(* IEC 61131-3 sources: veristc/veri-stc/tests/st-examples (part 4) *)

cond_a := LimitHigh(raw_110_a, 130);
cond_a := cond_a AND quality_a;
cond_a := cond_a AND (NOT bypass_a);
input_valid_a := InputValid(raw_110_a, 0, 1000);
cond_a := cond_a AND input_valid_a;
IF NOT input_valid_a THEN
    channel_fault_a := channel_fault_a + 1;
END_IF;
cond_b := LimitHigh(raw_110_b, 130);
cond_b := cond_b AND quality_b;
cond_b := cond_b AND (NOT bypass_b);
input_valid_b := InputValid(raw_110_b, 0, 1000);
cond_b := cond_b AND input_valid_b;
IF NOT input_valid_b THEN
    channel_fault_b := channel_fault_b + 1;
END_IF;
cond_c := LimitHigh(raw_110_c, 130);
cond_c := cond_c AND quality_c;
cond_c := cond_c AND (NOT bypass_c);
input_valid_c := InputValid(raw_110_c, 0, 1000);
cond_c := cond_c AND input_valid_c;
IF NOT input_valid_c THEN
    channel_fault_c := channel_fault_c + 1;
END_IF;
cond_d := LimitHigh(raw_110_d, 130);
cond_d := cond_d AND quality_d;
cond_d := cond_d AND (NOT bypass_d);
input_valid_d := InputValid(raw_110_d, 0, 1000);
cond_d := cond_d AND input_valid_d;
IF NOT input_valid_d THEN
    channel_fault_d := channel_fault_d + 1;
END_IF;
vote_ok := TwoOfFour(cond_a, cond_b, cond_c, cond_d);
IF cond_a <> cond_b THEN
    diagnosis_count := diagnosis_count + 1;
END_IF;
IF cond_c <> cond_d THEN
    diagnosis_count := diagnosis_count + 1;
END_IF;
IF NOT vote_ok THEN
    diagnosis_count := diagnosis_count + 1;
END_IF;
latch_a_110 := RS_Next(vote_ok, train_a_reset, latch_a_110);
IF latch_a_110 AND (NOT train_a_inhibit) THEN
    mask_a_13 := mask_a_13 + 64;
    trip_a := 0 < 1;
    scram_a := 0 < 1;
    breaker_a := 0 > 1;
    mfw_a := 0 < 1;
    alarm_a := 0 < 1;
END_IF;
latch_b_110 := RS_Next(vote_ok, train_b_reset, latch_b_110);
IF latch_b_110 AND (NOT train_b_inhibit) THEN
    mask_b_13 := mask_b_13 + 64;
    trip_b := 0 < 1;
    scram_b := 0 < 1;
    breaker_b := 0 > 1;
    mfw_b := 0 < 1;
    alarm_b := 0 < 1;
END_IF;
IF (raw_110_a > 130) AND (NOT cond_a) THEN
    channel_fault_a := channel_fault_a + 1;
END_IF;
IF (raw_110_b > 130) AND (NOT cond_b) THEN
    channel_fault_b := channel_fault_b + 1;
END_IF;
IF (raw_110_c > 130) AND (NOT cond_c) THEN
    channel_fault_c := channel_fault_c + 1;
END_IF;
IF (raw_110_d > 130) AND (NOT cond_d) THEN
    channel_fault_d := channel_fault_d + 1;
END_IF;
IF vote_ok AND train_a_inhibit THEN
    diagnosis_count := diagnosis_count + 1;
END_IF;
IF vote_ok AND train_b_inhibit THEN
    diagnosis_count := diagnosis_count + 1;
END_IF;

cond_a := LimitHigh(raw_111_a, 131);
cond_a := cond_a AND quality_a;
cond_a := cond_a AND (NOT bypass_a);
input_valid_a := InputValid(raw_111_a, 0, 1000);
cond_a := cond_a AND input_valid_a;
IF NOT input_valid_a THEN
    channel_fault_a := channel_fault_a + 1;
END_IF;
cond_b := LimitHigh(raw_111_b, 131);
cond_b := cond_b AND quality_b;
cond_b := cond_b AND (NOT bypass_b);
input_valid_b := InputValid(raw_111_b, 0, 1000);
cond_b := cond_b AND input_valid_b;
IF NOT input_valid_b THEN
    channel_fault_b := channel_fault_b + 1;
END_IF;
cond_c := LimitHigh(raw_111_c, 131);
cond_c := cond_c AND quality_c;
cond_c := cond_c AND (NOT bypass_c);
input_valid_c := InputValid(raw_111_c, 0, 1000);
cond_c := cond_c AND input_valid_c;
IF NOT input_valid_c THEN
    channel_fault_c := channel_fault_c + 1;
END_IF;
cond_d := LimitHigh(raw_111_d, 131);
cond_d := cond_d AND quality_d;
cond_d := cond_d AND (NOT bypass_d);
input_valid_d := InputValid(raw_111_d, 0, 1000);
cond_d := cond_d AND input_valid_d;
IF NOT input_valid_d THEN
    channel_fault_d := channel_fault_d + 1;
END_IF;
vote_ok := TwoOfFour(cond_a, cond_b, cond_c, cond_d);
IF cond_a <> cond_b THEN
    diagnosis_count := diagnosis_count + 1;
END_IF;
IF cond_c <> cond_d THEN
    diagnosis_count := diagnosis_count + 1;
END_IF;
IF NOT vote_ok THEN
    diagnosis_count := diagnosis_count + 1;
END_IF;
latch_a_111 := RS_Next(vote_ok, train_a_reset, latch_a_111);
IF latch_a_111 AND (NOT train_a_inhibit) THEN
    mask_a_13 := mask_a_13 + 128;
    trip_a := 0 < 1;
    scram_a := 0 < 1;
    breaker_a := 0 > 1;
    afw_a := 0 < 1;
    alarm_a := 0 < 1;
END_IF;
latch_b_111 := RS_Next(vote_ok, train_b_reset, latch_b_111);
IF latch_b_111 AND (NOT train_b_inhibit) THEN
    mask_b_13 := mask_b_13 + 128;
    trip_b := 0 < 1;
    scram_b := 0 < 1;
    breaker_b := 0 > 1;
    afw_b := 0 < 1;
    alarm_b := 0 < 1;
END_IF;
IF (raw_111_a > 131) AND (NOT cond_a) THEN
    channel_fault_a := channel_fault_a + 1;
END_IF;
IF (raw_111_b > 131) AND (NOT cond_b) THEN
    channel_fault_b := channel_fault_b + 1;
END_IF;
IF (raw_111_c > 131) AND (NOT cond_c) THEN
    channel_fault_c := channel_fault_c + 1;
END_IF;
IF (raw_111_d > 131) AND (NOT cond_d) THEN
    channel_fault_d := channel_fault_d + 1;
END_IF;
IF vote_ok AND train_a_inhibit THEN
    diagnosis_count := diagnosis_count + 1;
END_IF;
IF vote_ok AND train_b_inhibit THEN
    diagnosis_count := diagnosis_count + 1;
END_IF;

cond_a := LimitHigh(raw_112_a, 132);
cond_a := cond_a AND quality_a;
cond_a := cond_a AND (NOT bypass_a);
input_valid_a := InputValid(raw_112_a, 0, 1000);
cond_a := cond_a AND input_valid_a;
IF NOT input_valid_a THEN
    channel_fault_a := channel_fault_a + 1;
END_IF;
cond_b := LimitHigh(raw_112_b, 132);
cond_b := cond_b AND quality_b;
cond_b := cond_b AND (NOT bypass_b);
input_valid_b := InputValid(raw_112_b, 0, 1000);
cond_b := cond_b AND input_valid_b;
IF NOT input_valid_b THEN
    channel_fault_b := channel_fault_b + 1;
END_IF;
cond_c := LimitHigh(raw_112_c, 132);
cond_c := cond_c AND quality_c;
cond_c := cond_c AND (NOT bypass_c);
input_valid_c := InputValid(raw_112_c, 0, 1000);
cond_c := cond_c AND input_valid_c;
IF NOT input_valid_c THEN
    channel_fault_c := channel_fault_c + 1;
END_IF;
cond_d := LimitHigh(raw_112_d, 132);
cond_d := cond_d AND quality_d;
cond_d := cond_d AND (NOT bypass_d);
input_valid_d := InputValid(raw_112_d, 0, 1000);
cond_d := cond_d AND input_valid_d;
IF NOT input_valid_d THEN
    channel_fault_d := channel_fault_d + 1;
END_IF;
vote_ok := TwoOfFour(cond_a, cond_b, cond_c, cond_d);
IF cond_a <> cond_b THEN
    diagnosis_count := diagnosis_count + 1;
END_IF;
IF cond_c <> cond_d THEN
    diagnosis_count := diagnosis_count + 1;
END_IF;
IF NOT vote_ok THEN
    diagnosis_count := diagnosis_count + 1;
END_IF;
latch_a_112 := RS_Next(vote_ok, train_a_reset, latch_a_112);
IF latch_a_112 AND (NOT train_a_inhibit) THEN
    mask_a_14 := mask_a_14 + 1;
    trip_a := 0 < 1;
    scram_a := 0 < 1;
    breaker_a := 0 > 1;
    si_a := 0 < 1;
    alarm_a := 0 < 1;
END_IF;
latch_b_112 := RS_Next(vote_ok, train_b_reset, latch_b_112);
IF latch_b_112 AND (NOT train_b_inhibit) THEN
    mask_b_14 := mask_b_14 + 1;
    trip_b := 0 < 1;
    scram_b := 0 < 1;
    breaker_b := 0 > 1;
    si_b := 0 < 1;
    alarm_b := 0 < 1;
END_IF;
IF (raw_112_a > 132) AND (NOT cond_a) THEN
    channel_fault_a := channel_fault_a + 1;
END_IF;
IF (raw_112_b > 132) AND (NOT cond_b) THEN
    channel_fault_b := channel_fault_b + 1;
END_IF;
IF (raw_112_c > 132) AND (NOT cond_c) THEN
    channel_fault_c := channel_fault_c + 1;
END_IF;
IF (raw_112_d > 132) AND (NOT cond_d) THEN
    channel_fault_d := channel_fault_d + 1;
END_IF;
IF vote_ok AND train_a_inhibit THEN
    diagnosis_count := diagnosis_count + 1;
END_IF;
IF vote_ok AND train_b_inhibit THEN
    diagnosis_count := diagnosis_count + 1;
END_IF;

cond_a := LimitHigh(raw_113_a, 133);
cond_a := cond_a AND quality_a;
cond_a := cond_a AND (NOT bypass_a);
input_valid_a := InputValid(raw_113_a, 0, 1000);
cond_a := cond_a AND input_valid_a;
IF NOT input_valid_a THEN
    channel_fault_a := channel_fault_a + 1;
END_IF;
cond_b := LimitHigh(raw_113_b, 133);
cond_b := cond_b AND quality_b;
cond_b := cond_b AND (NOT bypass_b);
input_valid_b := InputValid(raw_113_b, 0, 1000);
cond_b := cond_b AND input_valid_b;
IF NOT input_valid_b THEN
    channel_fault_b := channel_fault_b + 1;
END_IF;
cond_c := LimitHigh(raw_113_c, 133);
cond_c := cond_c AND quality_c;
cond_c := cond_c AND (NOT bypass_c);
input_valid_c := InputValid(raw_113_c, 0, 1000);
cond_c := cond_c AND input_valid_c;
IF NOT input_valid_c THEN
    channel_fault_c := channel_fault_c + 1;
END_IF;
cond_d := LimitHigh(raw_113_d, 133);
cond_d := cond_d AND quality_d;
cond_d := cond_d AND (NOT bypass_d);
input_valid_d := InputValid(raw_113_d, 0, 1000);
cond_d := cond_d AND input_valid_d;
IF NOT input_valid_d THEN
    channel_fault_d := channel_fault_d + 1;
END_IF;
vote_ok := TwoOfFour(cond_a, cond_b, cond_c, cond_d);
IF cond_a <> cond_b THEN
    diagnosis_count := diagnosis_count + 1;
END_IF;
IF cond_c <> cond_d THEN
    diagnosis_count := diagnosis_count + 1;
END_IF;
IF NOT vote_ok THEN
    diagnosis_count := diagnosis_count + 1;
END_IF;
latch_a_113 := RS_Next(vote_ok, train_a_reset, latch_a_113);
IF latch_a_113 AND (NOT train_a_inhibit) THEN
    mask_a_14 := mask_a_14 + 2;
    trip_a := 0 < 1;
    scram_a := 0 < 1;
    breaker_a := 0 > 1;
    ci_a := 0 < 1;
    alarm_a := 0 < 1;
END_IF;
latch_b_113 := RS_Next(vote_ok, train_b_reset, latch_b_113);
IF latch_b_113 AND (NOT train_b_inhibit) THEN
    mask_b_14 := mask_b_14 + 2;
    trip_b := 0 < 1;
    scram_b := 0 < 1;
    breaker_b := 0 > 1;
    ci_b := 0 < 1;
    alarm_b := 0 < 1;
END_IF;
IF (raw_113_a > 133) AND (NOT cond_a) THEN
    channel_fault_a := channel_fault_a + 1;
END_IF;
IF (raw_113_b > 133) AND (NOT cond_b) THEN
    channel_fault_b := channel_fault_b + 1;
END_IF;
IF (raw_113_c > 133) AND (NOT cond_c) THEN
    channel_fault_c := channel_fault_c + 1;
END_IF;
IF (raw_113_d > 133) AND (NOT cond_d) THEN
    channel_fault_d := channel_fault_d + 1;
END_IF;
IF vote_ok AND train_a_inhibit THEN
    diagnosis_count := diagnosis_count + 1;
END_IF;
IF vote_ok AND train_b_inhibit THEN
    diagnosis_count := diagnosis_count + 1;
END_IF;

cond_a := LimitHigh(raw_114_a, 134);
cond_a := cond_a AND quality_a;
cond_a := cond_a AND (NOT bypass_a);
input_valid_a := InputValid(raw_114_a, 0, 1000);
cond_a := cond_a AND input_valid_a;
IF NOT input_valid_a THEN
    channel_fault_a := channel_fault_a + 1;
END_IF;
cond_b := LimitHigh(raw_114_b, 134);
cond_b := cond_b AND quality_b;
cond_b := cond_b AND (NOT bypass_b);
input_valid_b := InputValid(raw_114_b, 0, 1000);
cond_b := cond_b AND input_valid_b;
IF NOT input_valid_b THEN
    channel_fault_b := channel_fault_b + 1;
END_IF;
cond_c := LimitHigh(raw_114_c, 134);
cond_c := cond_c AND quality_c;
cond_c := cond_c AND (NOT bypass_c);
input_valid_c := InputValid(raw_114_c, 0, 1000);
cond_c := cond_c AND input_valid_c;
IF NOT input_valid_c THEN
    channel_fault_c := channel_fault_c + 1;
END_IF;
cond_d := LimitHigh(raw_114_d, 134);
cond_d := cond_d AND quality_d;
cond_d := cond_d AND (NOT bypass_d);
input_valid_d := InputValid(raw_114_d, 0, 1000);
cond_d := cond_d AND input_valid_d;
IF NOT input_valid_d THEN
    channel_fault_d := channel_fault_d + 1;
END_IF;
vote_ok := TwoOfFour(cond_a, cond_b, cond_c, cond_d);
IF cond_a <> cond_b THEN
    diagnosis_count := diagnosis_count + 1;
END_IF;
IF cond_c <> cond_d THEN
    diagnosis_count := diagnosis_count + 1;
END_IF;
IF NOT vote_ok THEN
    diagnosis_count := diagnosis_count + 1;
END_IF;
latch_a_114 := RS_Next(vote_ok, train_a_reset, latch_a_114);
IF latch_a_114 AND (NOT train_a_inhibit) THEN
    mask_a_14 := mask_a_14 + 4;
    trip_a := 0 < 1;
    scram_a := 0 < 1;
    breaker_a := 0 > 1;
    mfw_a := 0 < 1;
    alarm_a := 0 < 1;
END_IF;
latch_b_114 := RS_Next(vote_ok, train_b_reset, latch_b_114);
IF latch_b_114 AND (NOT train_b_inhibit) THEN
    mask_b_14 := mask_b_14 + 4;
    trip_b := 0 < 1;
    scram_b := 0 < 1;
    breaker_b := 0 > 1;
    mfw_b := 0 < 1;
    alarm_b := 0 < 1;
END_IF;
IF (raw_114_a > 134) AND (NOT cond_a) THEN
    channel_fault_a := channel_fault_a + 1;
END_IF;
IF (raw_114_b > 134) AND (NOT cond_b) THEN
    channel_fault_b := channel_fault_b + 1;
END_IF;
IF (raw_114_c > 134) AND (NOT cond_c) THEN
    channel_fault_c := channel_fault_c + 1;
END_IF;
IF (raw_114_d > 134) AND (NOT cond_d) THEN
    channel_fault_d := channel_fault_d + 1;
END_IF;
IF vote_ok AND train_a_inhibit THEN
    diagnosis_count := diagnosis_count + 1;
END_IF;
IF vote_ok AND train_b_inhibit THEN
    diagnosis_count := diagnosis_count + 1;
END_IF;

cond_a := LimitHigh(raw_115_a, 135);
cond_a := cond_a AND quality_a;
cond_a := cond_a AND (NOT bypass_a);
input_valid_a := InputValid(raw_115_a, 0, 1000);
cond_a := cond_a AND input_valid_a;
IF NOT input_valid_a THEN
    channel_fault_a := channel_fault_a + 1;
END_IF;
cond_b := LimitHigh(raw_115_b, 135);
cond_b := cond_b AND quality_b;
cond_b := cond_b AND (NOT bypass_b);
input_valid_b := InputValid(raw_115_b, 0, 1000);
cond_b := cond_b AND input_valid_b;
IF NOT input_valid_b THEN
    channel_fault_b := channel_fault_b + 1;
END_IF;
cond_c := LimitHigh(raw_115_c, 135);
cond_c := cond_c AND quality_c;
cond_c := cond_c AND (NOT bypass_c);
input_valid_c := InputValid(raw_115_c, 0, 1000);
cond_c := cond_c AND input_valid_c;
IF NOT input_valid_c THEN
    channel_fault_c := channel_fault_c + 1;
END_IF;
cond_d := LimitHigh(raw_115_d, 135);
cond_d := cond_d AND quality_d;
cond_d := cond_d AND (NOT bypass_d);
input_valid_d := InputValid(raw_115_d, 0, 1000);
cond_d := cond_d AND input_valid_d;
IF NOT input_valid_d THEN
    channel_fault_d := channel_fault_d + 1;
END_IF;
vote_ok := TwoOfFour(cond_a, cond_b, cond_c, cond_d);
IF cond_a <> cond_b THEN
    diagnosis_count := diagnosis_count + 1;
END_IF;
IF cond_c <> cond_d THEN
    diagnosis_count := diagnosis_count + 1;
END_IF;
IF NOT vote_ok THEN
    diagnosis_count := diagnosis_count + 1;
END_IF;
latch_a_115 := RS_Next(vote_ok, train_a_reset, latch_a_115);
IF latch_a_115 AND (NOT train_a_inhibit) THEN
    mask_a_14 := mask_a_14 + 8;
    trip_a := 0 < 1;
    scram_a := 0 < 1;
    breaker_a := 0 > 1;
    afw_a := 0 < 1;
    alarm_a := 0 < 1;
END_IF;
latch_b_115 := RS_Next(vote_ok, train_b_reset, latch_b_115);
IF latch_b_115 AND (NOT train_b_inhibit) THEN
    mask_b_14 := mask_b_14 + 8;
    trip_b := 0 < 1;
    scram_b := 0 < 1;
    breaker_b := 0 > 1;
    afw_b := 0 < 1;
    alarm_b := 0 < 1;
END_IF;
IF (raw_115_a > 135) AND (NOT cond_a) THEN
    channel_fault_a := channel_fault_a + 1;
END_IF;
IF (raw_115_b > 135) AND (NOT cond_b) THEN
    channel_fault_b := channel_fault_b + 1;
END_IF;
IF (raw_115_c > 135) AND (NOT cond_c) THEN
    channel_fault_c := channel_fault_c + 1;
END_IF;
IF (raw_115_d > 135) AND (NOT cond_d) THEN
    channel_fault_d := channel_fault_d + 1;
END_IF;
IF vote_ok AND train_a_inhibit THEN
    diagnosis_count := diagnosis_count + 1;
END_IF;
IF vote_ok AND train_b_inhibit THEN
    diagnosis_count := diagnosis_count + 1;
END_IF;

cond_a := LimitHigh(raw_116_a, 136);
cond_a := cond_a AND quality_a;
cond_a := cond_a AND (NOT bypass_a);
input_valid_a := InputValid(raw_116_a, 0, 1000);
cond_a := cond_a AND input_valid_a;
IF NOT input_valid_a THEN
    channel_fault_a := channel_fault_a + 1;
END_IF;
cond_b := LimitHigh(raw_116_b, 136);
cond_b := cond_b AND quality_b;
cond_b := cond_b AND (NOT bypass_b);
input_valid_b := InputValid(raw_116_b, 0, 1000);
cond_b := cond_b AND input_valid_b;
IF NOT input_valid_b THEN
    channel_fault_b := channel_fault_b + 1;
END_IF;
cond_c := LimitHigh(raw_116_c, 136);
cond_c := cond_c AND quality_c;
cond_c := cond_c AND (NOT bypass_c);
input_valid_c := InputValid(raw_116_c, 0, 1000);
cond_c := cond_c AND input_valid_c;
IF NOT input_valid_c THEN
    channel_fault_c := channel_fault_c + 1;
END_IF;
cond_d := LimitHigh(raw_116_d, 136);
cond_d := cond_d AND quality_d;
cond_d := cond_d AND (NOT bypass_d);
input_valid_d := InputValid(raw_116_d, 0, 1000);
cond_d := cond_d AND input_valid_d;
IF NOT input_valid_d THEN
    channel_fault_d := channel_fault_d + 1;
END_IF;
vote_ok := TwoOfFour(cond_a, cond_b, cond_c, cond_d);
IF cond_a <> cond_b THEN
    diagnosis_count := diagnosis_count + 1;
END_IF;
IF cond_c <> cond_d THEN
    diagnosis_count := diagnosis_count + 1;
END_IF;
IF NOT vote_ok THEN
    diagnosis_count := diagnosis_count + 1;
END_IF;
latch_a_116 := RS_Next(vote_ok, train_a_reset, latch_a_116);
IF latch_a_116 AND (NOT train_a_inhibit) THEN
    mask_a_14 := mask_a_14 + 16;
    trip_a := 0 < 1;
    scram_a := 0 < 1;
    breaker_a := 0 > 1;
    si_a := 0 < 1;
    alarm_a := 0 < 1;
END_IF;
latch_b_116 := RS_Next(vote_ok, train_b_reset, latch_b_116);
IF latch_b_116 AND (NOT train_b_inhibit) THEN
    mask_b_14 := mask_b_14 + 16;
    trip_b := 0 < 1;
    scram_b := 0 < 1;
    breaker_b := 0 > 1;
    si_b := 0 < 1;
    alarm_b := 0 < 1;
END_IF;
IF (raw_116_a > 136) AND (NOT cond_a) THEN
    channel_fault_a := channel_fault_a + 1;
END_IF;
IF (raw_116_b > 136) AND (NOT cond_b) THEN
    channel_fault_b := channel_fault_b + 1;
END_IF;
IF (raw_116_c > 136) AND (NOT cond_c) THEN
    channel_fault_c := channel_fault_c + 1;
END_IF;
IF (raw_116_d > 136) AND (NOT cond_d) THEN
    channel_fault_d := channel_fault_d + 1;
END_IF;
IF vote_ok AND train_a_inhibit THEN
    diagnosis_count := diagnosis_count + 1;
END_IF;
IF vote_ok AND train_b_inhibit THEN
    diagnosis_count := diagnosis_count + 1;
END_IF;

cond_a := LimitHigh(raw_117_a, 137);
cond_a := cond_a AND quality_a;
cond_a := cond_a AND (NOT bypass_a);
input_valid_a := InputValid(raw_117_a, 0, 1000);
cond_a := cond_a AND input_valid_a;
IF NOT input_valid_a THEN
    channel_fault_a := channel_fault_a + 1;
END_IF;
cond_b := LimitHigh(raw_117_b, 137);
cond_b := cond_b AND quality_b;
cond_b := cond_b AND (NOT bypass_b);
input_valid_b := InputValid(raw_117_b, 0, 1000);
cond_b := cond_b AND input_valid_b;
IF NOT input_valid_b THEN
    channel_fault_b := channel_fault_b + 1;
END_IF;
cond_c := LimitHigh(raw_117_c, 137);
cond_c := cond_c AND quality_c;
cond_c := cond_c AND (NOT bypass_c);
input_valid_c := InputValid(raw_117_c, 0, 1000);
cond_c := cond_c AND input_valid_c;
IF NOT input_valid_c THEN
    channel_fault_c := channel_fault_c + 1;
END_IF;
cond_d := LimitHigh(raw_117_d, 137);
cond_d := cond_d AND quality_d;
cond_d := cond_d AND (NOT bypass_d);
input_valid_d := InputValid(raw_117_d, 0, 1000);
cond_d := cond_d AND input_valid_d;
IF NOT input_valid_d THEN
    channel_fault_d := channel_fault_d + 1;
END_IF;
vote_ok := TwoOfFour(cond_a, cond_b, cond_c, cond_d);
IF cond_a <> cond_b THEN
    diagnosis_count := diagnosis_count + 1;
END_IF;
IF cond_c <> cond_d THEN
    diagnosis_count := diagnosis_count + 1;
END_IF;
IF NOT vote_ok THEN
    diagnosis_count := diagnosis_count + 1;
END_IF;
latch_a_117 := RS_Next(vote_ok, train_a_reset, latch_a_117);
IF latch_a_117 AND (NOT train_a_inhibit) THEN
    mask_a_14 := mask_a_14 + 32;
    trip_a := 0 < 1;
    scram_a := 0 < 1;
    breaker_a := 0 > 1;
    ci_a := 0 < 1;
    alarm_a := 0 < 1;
END_IF;
latch_b_117 := RS_Next(vote_ok, train_b_reset, latch_b_117);
IF latch_b_117 AND (NOT train_b_inhibit) THEN
    mask_b_14 := mask_b_14 + 32;
    trip_b := 0 < 1;
    scram_b := 0 < 1;
    breaker_b := 0 > 1;
    ci_b := 0 < 1;
    alarm_b := 0 < 1;
END_IF;
IF (raw_117_a > 137) AND (NOT cond_a) THEN
    channel_fault_a := channel_fault_a + 1;
END_IF;
IF (raw_117_b > 137) AND (NOT cond_b) THEN
    channel_fault_b := channel_fault_b + 1;
END_IF;
IF (raw_117_c > 137) AND (NOT cond_c) THEN
    channel_fault_c := channel_fault_c + 1;
END_IF;
IF (raw_117_d > 137) AND (NOT cond_d) THEN
    channel_fault_d := channel_fault_d + 1;
END_IF;
IF vote_ok AND train_a_inhibit THEN
    diagnosis_count := diagnosis_count + 1;
END_IF;
IF vote_ok AND train_b_inhibit THEN
    diagnosis_count := diagnosis_count + 1;
END_IF;

cond_a := LimitHigh(raw_118_a, 138);
cond_a := cond_a AND quality_a;
cond_a := cond_a AND (NOT bypass_a);
input_valid_a := InputValid(raw_118_a, 0, 1000);
cond_a := cond_a AND input_valid_a;
IF NOT input_valid_a THEN
    channel_fault_a := channel_fault_a + 1;
END_IF;
cond_b := LimitHigh(raw_118_b, 138);
cond_b := cond_b AND quality_b;
cond_b := cond_b AND (NOT bypass_b);
input_valid_b := InputValid(raw_118_b, 0, 1000);
cond_b := cond_b AND input_valid_b;
IF NOT input_valid_b THEN
    channel_fault_b := channel_fault_b + 1;
END_IF;
cond_c := LimitHigh(raw_118_c, 138);
cond_c := cond_c AND quality_c;
cond_c := cond_c AND (NOT bypass_c);
input_valid_c := InputValid(raw_118_c, 0, 1000);
cond_c := cond_c AND input_valid_c;
IF NOT input_valid_c THEN
    channel_fault_c := channel_fault_c + 1;
END_IF;
cond_d := LimitHigh(raw_118_d, 138);
cond_d := cond_d AND quality_d;
cond_d := cond_d AND (NOT bypass_d);
input_valid_d := InputValid(raw_118_d, 0, 1000);
cond_d := cond_d AND input_valid_d;
IF NOT input_valid_d THEN
    channel_fault_d := channel_fault_d + 1;
END_IF;
vote_ok := TwoOfFour(cond_a, cond_b, cond_c, cond_d);
IF cond_a <> cond_b THEN
    diagnosis_count := diagnosis_count + 1;
END_IF;
IF cond_c <> cond_d THEN
    diagnosis_count := diagnosis_count + 1;
END_IF;
IF NOT vote_ok THEN
    diagnosis_count := diagnosis_count + 1;
END_IF;
latch_a_118 := RS_Next(vote_ok, train_a_reset, latch_a_118);
IF latch_a_118 AND (NOT train_a_inhibit) THEN
    mask_a_14 := mask_a_14 + 64;
    trip_a := 0 < 1;
    scram_a := 0 < 1;
    breaker_a := 0 > 1;
    mfw_a := 0 < 1;
    alarm_a := 0 < 1;
END_IF;
latch_b_118 := RS_Next(vote_ok, train_b_reset, latch_b_118);
IF latch_b_118 AND (NOT train_b_inhibit) THEN
    mask_b_14 := mask_b_14 + 64;
    trip_b := 0 < 1;
    scram_b := 0 < 1;
    breaker_b := 0 > 1;
    mfw_b := 0 < 1;
    alarm_b := 0 < 1;
END_IF;
IF (raw_118_a > 138) AND (NOT cond_a) THEN
    channel_fault_a := channel_fault_a + 1;
END_IF;
IF (raw_118_b > 138) AND (NOT cond_b) THEN
    channel_fault_b := channel_fault_b + 1;
END_IF;
IF (raw_118_c > 138) AND (NOT cond_c) THEN
    channel_fault_c := channel_fault_c + 1;
END_IF;
IF (raw_118_d > 138) AND (NOT cond_d) THEN
    channel_fault_d := channel_fault_d + 1;
END_IF;
IF vote_ok AND train_a_inhibit THEN
    diagnosis_count := diagnosis_count + 1;
END_IF;
IF vote_ok AND train_b_inhibit THEN
    diagnosis_count := diagnosis_count + 1;
END_IF;

cond_a := LimitHigh(raw_119_a, 139);
cond_a := cond_a AND quality_a;
cond_a := cond_a AND (NOT bypass_a);
input_valid_a := InputValid(raw_119_a, 0, 1000);
cond_a := cond_a AND input_valid_a;
IF NOT input_valid_a THEN
    channel_fault_a := channel_fault_a + 1;
END_IF;
cond_b := LimitHigh(raw_119_b, 139);
cond_b := cond_b AND quality_b;
cond_b := cond_b AND (NOT bypass_b);
input_valid_b := InputValid(raw_119_b, 0, 1000);
cond_b := cond_b AND input_valid_b;
IF NOT input_valid_b THEN
    channel_fault_b := channel_fault_b + 1;
END_IF;
cond_c := LimitHigh(raw_119_c, 139);
cond_c := cond_c AND quality_c;
cond_c := cond_c AND (NOT bypass_c);
input_valid_c := InputValid(raw_119_c, 0, 1000);
cond_c := cond_c AND input_valid_c;
IF NOT input_valid_c THEN
    channel_fault_c := channel_fault_c + 1;
END_IF;
cond_d := LimitHigh(raw_119_d, 139);
cond_d := cond_d AND quality_d;
cond_d := cond_d AND (NOT bypass_d);
input_valid_d := InputValid(raw_119_d, 0, 1000);
cond_d := cond_d AND input_valid_d;
IF NOT input_valid_d THEN
    channel_fault_d := channel_fault_d + 1;
END_IF;
vote_ok := TwoOfFour(cond_a, cond_b, cond_c, cond_d);
IF cond_a <> cond_b THEN
    diagnosis_count := diagnosis_count + 1;
END_IF;
IF cond_c <> cond_d THEN
    diagnosis_count := diagnosis_count + 1;
END_IF;
IF NOT vote_ok THEN
    diagnosis_count := diagnosis_count + 1;
END_IF;
latch_a_119 := RS_Next(vote_ok, train_a_reset, latch_a_119);
IF latch_a_119 AND (NOT train_a_inhibit) THEN
    mask_a_14 := mask_a_14 + 128;
    trip_a := 0 < 1;
    scram_a := 0 < 1;
    breaker_a := 0 > 1;
    afw_a := 0 < 1;
    alarm_a := 0 < 1;
END_IF;
latch_b_119 := RS_Next(vote_ok, train_b_reset, latch_b_119);
IF latch_b_119 AND (NOT train_b_inhibit) THEN
    mask_b_14 := mask_b_14 + 128;
    trip_b := 0 < 1;
    scram_b := 0 < 1;
    breaker_b := 0 > 1;
    afw_b := 0 < 1;
    alarm_b := 0 < 1;
END_IF;
IF (raw_119_a > 139) AND (NOT cond_a) THEN
    channel_fault_a := channel_fault_a + 1;
END_IF;
IF (raw_119_b > 139) AND (NOT cond_b) THEN
    channel_fault_b := channel_fault_b + 1;
END_IF;
IF (raw_119_c > 139) AND (NOT cond_c) THEN
    channel_fault_c := channel_fault_c + 1;
END_IF;
IF (raw_119_d > 139) AND (NOT cond_d) THEN
    channel_fault_d := channel_fault_d + 1;
END_IF;
IF vote_ok AND train_a_inhibit THEN
    diagnosis_count := diagnosis_count + 1;
END_IF;
IF vote_ok AND train_b_inhibit THEN
    diagnosis_count := diagnosis_count + 1;
END_IF;

cond_a := LimitHigh(raw_120_a, 100);
cond_a := cond_a AND quality_a;
cond_a := cond_a AND (NOT bypass_a);
input_valid_a := InputValid(raw_120_a, 0, 1000);
cond_a := cond_a AND input_valid_a;
IF NOT input_valid_a THEN
    channel_fault_a := channel_fault_a + 1;
END_IF;
cond_b := LimitHigh(raw_120_b, 100);
cond_b := cond_b AND quality_b;
cond_b := cond_b AND (NOT bypass_b);
input_valid_b := InputValid(raw_120_b, 0, 1000);
cond_b := cond_b AND input_valid_b;
IF NOT input_valid_b THEN
    channel_fault_b := channel_fault_b + 1;
END_IF;
cond_c := LimitHigh(raw_120_c, 100);
cond_c := cond_c AND quality_c;
cond_c := cond_c AND (NOT bypass_c);
input_valid_c := InputValid(raw_120_c, 0, 1000);
cond_c := cond_c AND input_valid_c;
IF NOT input_valid_c THEN
    channel_fault_c := channel_fault_c + 1;
END_IF;
cond_d := LimitHigh(raw_120_d, 100);
cond_d := cond_d AND quality_d;
cond_d := cond_d AND (NOT bypass_d);
input_valid_d := InputValid(raw_120_d, 0, 1000);
cond_d := cond_d AND input_valid_d;
IF NOT input_valid_d THEN
    channel_fault_d := channel_fault_d + 1;
END_IF;
vote_ok := TwoOfFour(cond_a, cond_b, cond_c, cond_d);
IF cond_a <> cond_b THEN
    diagnosis_count := diagnosis_count + 1;
END_IF;
IF cond_c <> cond_d THEN
    diagnosis_count := diagnosis_count + 1;
END_IF;
IF NOT vote_ok THEN
    diagnosis_count := diagnosis_count + 1;
END_IF;
latch_a_120 := RS_Next(vote_ok, train_a_reset, latch_a_120);
IF latch_a_120 AND (NOT train_a_inhibit) THEN
    mask_a_15 := mask_a_15 + 1;
    trip_a := 0 < 1;
    scram_a := 0 < 1;
    breaker_a := 0 > 1;
    si_a := 0 < 1;
    alarm_a := 0 < 1;
END_IF;
latch_b_120 := RS_Next(vote_ok, train_b_reset, latch_b_120);
IF latch_b_120 AND (NOT train_b_inhibit) THEN
    mask_b_15 := mask_b_15 + 1;
    trip_b := 0 < 1;
    scram_b := 0 < 1;
    breaker_b := 0 > 1;
    si_b := 0 < 1;
    alarm_b := 0 < 1;
END_IF;
IF (raw_120_a > 100) AND (NOT cond_a) THEN
    channel_fault_a := channel_fault_a + 1;
END_IF;
IF (raw_120_b > 100) AND (NOT cond_b) THEN
    channel_fault_b := channel_fault_b + 1;
END_IF;
IF (raw_120_c > 100) AND (NOT cond_c) THEN
    channel_fault_c := channel_fault_c + 1;
END_IF;
IF (raw_120_d > 100) AND (NOT cond_d) THEN
    channel_fault_d := channel_fault_d + 1;
END_IF;
IF vote_ok AND train_a_inhibit THEN
    diagnosis_count := diagnosis_count + 1;
END_IF;
IF vote_ok AND train_b_inhibit THEN
    diagnosis_count := diagnosis_count + 1;
END_IF;

cond_a := LimitHigh(raw_121_a, 101);
cond_a := cond_a AND quality_a;
cond_a := cond_a AND (NOT bypass_a);
input_valid_a := InputValid(raw_121_a, 0, 1000);
cond_a := cond_a AND input_valid_a;
IF NOT input_valid_a THEN
    channel_fault_a := channel_fault_a + 1;
END_IF;
cond_b := LimitHigh(raw_121_b, 101);
cond_b := cond_b AND quality_b;
cond_b := cond_b AND (NOT bypass_b);
input_valid_b := InputValid(raw_121_b, 0, 1000);
cond_b := cond_b AND input_valid_b;
IF NOT input_valid_b THEN
    channel_fault_b := channel_fault_b + 1;
END_IF;
cond_c := LimitHigh(raw_121_c, 101);
cond_c := cond_c AND quality_c;
cond_c := cond_c AND (NOT bypass_c);
input_valid_c := InputValid(raw_121_c, 0, 1000);
cond_c := cond_c AND input_valid_c;
IF NOT input_valid_c THEN
    channel_fault_c := channel_fault_c + 1;
END_IF;
cond_d := LimitHigh(raw_121_d, 101);
cond_d := cond_d AND quality_d;
cond_d := cond_d AND (NOT bypass_d);
input_valid_d := InputValid(raw_121_d, 0, 1000);
cond_d := cond_d AND input_valid_d;
IF NOT input_valid_d THEN
    channel_fault_d := channel_fault_d + 1;
END_IF;
vote_ok := TwoOfFour(cond_a, cond_b, cond_c, cond_d);
IF cond_a <> cond_b THEN
    diagnosis_count := diagnosis_count + 1;
END_IF;
IF cond_c <> cond_d THEN
    diagnosis_count := diagnosis_count + 1;
END_IF;
IF NOT vote_ok THEN
    diagnosis_count := diagnosis_count + 1;
END_IF;
latch_a_121 := RS_Next(vote_ok, train_a_reset, latch_a_121);
IF latch_a_121 AND (NOT train_a_inhibit) THEN
    mask_a_15 := mask_a_15 + 2;
    trip_a := 0 < 1;
    scram_a := 0 < 1;
    breaker_a := 0 > 1;
    ci_a := 0 < 1;
    alarm_a := 0 < 1;
END_IF;
latch_b_121 := RS_Next(vote_ok, train_b_reset, latch_b_121);
IF latch_b_121 AND (NOT train_b_inhibit) THEN
    mask_b_15 := mask_b_15 + 2;
    trip_b := 0 < 1;
    scram_b := 0 < 1;
    breaker_b := 0 > 1;
    ci_b := 0 < 1;
    alarm_b := 0 < 1;
END_IF;
IF (raw_121_a > 101) AND (NOT cond_a) THEN
    channel_fault_a := channel_fault_a + 1;
END_IF;
IF (raw_121_b > 101) AND (NOT cond_b) THEN
    channel_fault_b := channel_fault_b + 1;
END_IF;
IF (raw_121_c > 101) AND (NOT cond_c) THEN
    channel_fault_c := channel_fault_c + 1;
END_IF;
IF (raw_121_d > 101) AND (NOT cond_d) THEN
    channel_fault_d := channel_fault_d + 1;
END_IF;
IF vote_ok AND train_a_inhibit THEN
    diagnosis_count := diagnosis_count + 1;
END_IF;
IF vote_ok AND train_b_inhibit THEN
    diagnosis_count := diagnosis_count + 1;
END_IF;

cond_a := LimitHigh(raw_122_a, 102);
cond_a := cond_a AND quality_a;
cond_a := cond_a AND (NOT bypass_a);
input_valid_a := InputValid(raw_122_a, 0, 1000);
cond_a := cond_a AND input_valid_a;
IF NOT input_valid_a THEN
    channel_fault_a := channel_fault_a + 1;
END_IF;
cond_b := LimitHigh(raw_122_b, 102);
cond_b := cond_b AND quality_b;
cond_b := cond_b AND (NOT bypass_b);
input_valid_b := InputValid(raw_122_b, 0, 1000);
cond_b := cond_b AND input_valid_b;
IF NOT input_valid_b THEN
    channel_fault_b := channel_fault_b + 1;
END_IF;
cond_c := LimitHigh(raw_122_c, 102);
cond_c := cond_c AND quality_c;
cond_c := cond_c AND (NOT bypass_c);
input_valid_c := InputValid(raw_122_c, 0, 1000);
cond_c := cond_c AND input_valid_c;
IF NOT input_valid_c THEN
    channel_fault_c := channel_fault_c + 1;
END_IF;
cond_d := LimitHigh(raw_122_d, 102);
cond_d := cond_d AND quality_d;
cond_d := cond_d AND (NOT bypass_d);
input_valid_d := InputValid(raw_122_d, 0, 1000);
cond_d := cond_d AND input_valid_d;
IF NOT input_valid_d THEN
    channel_fault_d := channel_fault_d + 1;
END_IF;
vote_ok := TwoOfFour(cond_a, cond_b, cond_c, cond_d);
IF cond_a <> cond_b THEN
    diagnosis_count := diagnosis_count + 1;
END_IF;
IF cond_c <> cond_d THEN
    diagnosis_count := diagnosis_count + 1;
END_IF;
IF NOT vote_ok THEN
    diagnosis_count := diagnosis_count + 1;
END_IF;
latch_a_122 := RS_Next(vote_ok, train_a_reset, latch_a_122);
IF latch_a_122 AND (NOT train_a_inhibit) THEN
    mask_a_15 := mask_a_15 + 4;
    trip_a := 0 < 1;
    scram_a := 0 < 1;
    breaker_a := 0 > 1;
    mfw_a := 0 < 1;
    alarm_a := 0 < 1;
END_IF;
latch_b_122 := RS_Next(vote_ok, train_b_reset, latch_b_122);
IF latch_b_122 AND (NOT train_b_inhibit) THEN
    mask_b_15 := mask_b_15 + 4;
    trip_b := 0 < 1;
    scram_b := 0 < 1;
    breaker_b := 0 > 1;
    mfw_b := 0 < 1;
    alarm_b := 0 < 1;
END_IF;
IF (raw_122_a > 102) AND (NOT cond_a) THEN
    channel_fault_a := channel_fault_a + 1;
END_IF;
IF (raw_122_b > 102) AND (NOT cond_b) THEN
    channel_fault_b := channel_fault_b + 1;
END_IF;
IF (raw_122_c > 102) AND (NOT cond_c) THEN
    channel_fault_c := channel_fault_c + 1;
END_IF;
IF (raw_122_d > 102) AND (NOT cond_d) THEN
    channel_fault_d := channel_fault_d + 1;
END_IF;
IF vote_ok AND train_a_inhibit THEN
    diagnosis_count := diagnosis_count + 1;
END_IF;
IF vote_ok AND train_b_inhibit THEN
    diagnosis_count := diagnosis_count + 1;
END_IF;

cond_a := LimitHigh(raw_123_a, 103);
cond_a := cond_a AND quality_a;
cond_a := cond_a AND (NOT bypass_a);
input_valid_a := InputValid(raw_123_a, 0, 1000);
cond_a := cond_a AND input_valid_a;
IF NOT input_valid_a THEN
    channel_fault_a := channel_fault_a + 1;
END_IF;
cond_b := LimitHigh(raw_123_b, 103);
cond_b := cond_b AND quality_b;
cond_b := cond_b AND (NOT bypass_b);
input_valid_b := InputValid(raw_123_b, 0, 1000);
cond_b := cond_b AND input_valid_b;
IF NOT input_valid_b THEN
    channel_fault_b := channel_fault_b + 1;
END_IF;
cond_c := LimitHigh(raw_123_c, 103);
cond_c := cond_c AND quality_c;
cond_c := cond_c AND (NOT bypass_c);
input_valid_c := InputValid(raw_123_c, 0, 1000);
cond_c := cond_c AND input_valid_c;
IF NOT input_valid_c THEN
    channel_fault_c := channel_fault_c + 1;
END_IF;
cond_d := LimitHigh(raw_123_d, 103);
cond_d := cond_d AND quality_d;
cond_d := cond_d AND (NOT bypass_d);
input_valid_d := InputValid(raw_123_d, 0, 1000);
cond_d := cond_d AND input_valid_d;
IF NOT input_valid_d THEN
    channel_fault_d := channel_fault_d + 1;
END_IF;
vote_ok := TwoOfFour(cond_a, cond_b, cond_c, cond_d);
IF cond_a <> cond_b THEN
    diagnosis_count := diagnosis_count + 1;
END_IF;
IF cond_c <> cond_d THEN
    diagnosis_count := diagnosis_count + 1;
END_IF;
IF NOT vote_ok THEN
    diagnosis_count := diagnosis_count + 1;
END_IF;
latch_a_123 := RS_Next(vote_ok, train_a_reset, latch_a_123);
IF latch_a_123 AND (NOT train_a_inhibit) THEN
    mask_a_15 := mask_a_15 + 8;
    trip_a := 0 < 1;
    scram_a := 0 < 1;
    breaker_a := 0 > 1;
    afw_a := 0 < 1;
    alarm_a := 0 < 1;
END_IF;
latch_b_123 := RS_Next(vote_ok, train_b_reset, latch_b_123);
IF latch_b_123 AND (NOT train_b_inhibit) THEN
    mask_b_15 := mask_b_15 + 8;
    trip_b := 0 < 1;
    scram_b := 0 < 1;
    breaker_b := 0 > 1;
    afw_b := 0 < 1;
    alarm_b := 0 < 1;
END_IF;
IF (raw_123_a > 103) AND (NOT cond_a) THEN
    channel_fault_a := channel_fault_a + 1;
END_IF;
IF (raw_123_b > 103) AND (NOT cond_b) THEN
    channel_fault_b := channel_fault_b + 1;
END_IF;
IF (raw_123_c > 103) AND (NOT cond_c) THEN
    channel_fault_c := channel_fault_c + 1;
END_IF;
IF (raw_123_d > 103) AND (NOT cond_d) THEN
    channel_fault_d := channel_fault_d + 1;
END_IF;
IF vote_ok AND train_a_inhibit THEN
    diagnosis_count := diagnosis_count + 1;
END_IF;
IF vote_ok AND train_b_inhibit THEN
    diagnosis_count := diagnosis_count + 1;
END_IF;

cond_a := LimitHigh(raw_124_a, 104);
cond_a := cond_a AND quality_a;
cond_a := cond_a AND (NOT bypass_a);
input_valid_a := InputValid(raw_124_a, 0, 1000);
cond_a := cond_a AND input_valid_a;
IF NOT input_valid_a THEN
    channel_fault_a := channel_fault_a + 1;
END_IF;
cond_b := LimitHigh(raw_124_b, 104);
cond_b := cond_b AND quality_b;
cond_b := cond_b AND (NOT bypass_b);
input_valid_b := InputValid(raw_124_b, 0, 1000);
cond_b := cond_b AND input_valid_b;
IF NOT input_valid_b THEN
    channel_fault_b := channel_fault_b + 1;
END_IF;
cond_c := LimitHigh(raw_124_c, 104);
cond_c := cond_c AND quality_c;
cond_c := cond_c AND (NOT bypass_c);
input_valid_c := InputValid(raw_124_c, 0, 1000);
cond_c := cond_c AND input_valid_c;
IF NOT input_valid_c THEN
    channel_fault_c := channel_fault_c + 1;
END_IF;
cond_d := LimitHigh(raw_124_d, 104);
cond_d := cond_d AND quality_d;
cond_d := cond_d AND (NOT bypass_d);
input_valid_d := InputValid(raw_124_d, 0, 1000);
cond_d := cond_d AND input_valid_d;
IF NOT input_valid_d THEN
    channel_fault_d := channel_fault_d + 1;
END_IF;
vote_ok := TwoOfFour(cond_a, cond_b, cond_c, cond_d);
IF cond_a <> cond_b THEN
    diagnosis_count := diagnosis_count + 1;
END_IF;
IF cond_c <> cond_d THEN
    diagnosis_count := diagnosis_count + 1;
END_IF;
IF NOT vote_ok THEN
    diagnosis_count := diagnosis_count + 1;
END_IF;
latch_a_124 := RS_Next(vote_ok, train_a_reset, latch_a_124);
IF latch_a_124 AND (NOT train_a_inhibit) THEN
    mask_a_15 := mask_a_15 + 16;
    trip_a := 0 < 1;
    scram_a := 0 < 1;
    breaker_a := 0 > 1;
    si_a := 0 < 1;
    alarm_a := 0 < 1;
END_IF;
latch_b_124 := RS_Next(vote_ok, train_b_reset, latch_b_124);
IF latch_b_124 AND (NOT train_b_inhibit) THEN
    mask_b_15 := mask_b_15 + 16;
    trip_b := 0 < 1;
    scram_b := 0 < 1;
    breaker_b := 0 > 1;
    si_b := 0 < 1;
    alarm_b := 0 < 1;
END_IF;
IF (raw_124_a > 104) AND (NOT cond_a) THEN
    channel_fault_a := channel_fault_a + 1;
END_IF;
IF (raw_124_b > 104) AND (NOT cond_b) THEN
    channel_fault_b := channel_fault_b + 1;
END_IF;
IF (raw_124_c > 104) AND (NOT cond_c) THEN
    channel_fault_c := channel_fault_c + 1;
END_IF;
IF (raw_124_d > 104) AND (NOT cond_d) THEN
    channel_fault_d := channel_fault_d + 1;
END_IF;
IF vote_ok AND train_a_inhibit THEN
    diagnosis_count := diagnosis_count + 1;
END_IF;
IF vote_ok AND train_b_inhibit THEN
    diagnosis_count := diagnosis_count + 1;
END_IF;

cond_a := LimitHigh(raw_125_a, 105);
cond_a := cond_a AND quality_a;
cond_a := cond_a AND (NOT bypass_a);
input_valid_a := InputValid(raw_125_a, 0, 1000);
cond_a := cond_a AND input_valid_a;
IF NOT input_valid_a THEN
    channel_fault_a := channel_fault_a + 1;
END_IF;
cond_b := LimitHigh(raw_125_b, 105);
cond_b := cond_b AND quality_b;
cond_b := cond_b AND (NOT bypass_b);
input_valid_b := InputValid(raw_125_b, 0, 1000);
cond_b := cond_b AND input_valid_b;
IF NOT input_valid_b THEN
    channel_fault_b := channel_fault_b + 1;
END_IF;
cond_c := LimitHigh(raw_125_c, 105);
cond_c := cond_c AND quality_c;
cond_c := cond_c AND (NOT bypass_c);
input_valid_c := InputValid(raw_125_c, 0, 1000);
cond_c := cond_c AND input_valid_c;
IF NOT input_valid_c THEN
    channel_fault_c := channel_fault_c + 1;
END_IF;
cond_d := LimitHigh(raw_125_d, 105);
cond_d := cond_d AND quality_d;
cond_d := cond_d AND (NOT bypass_d);
input_valid_d := InputValid(raw_125_d, 0, 1000);
cond_d := cond_d AND input_valid_d;
IF NOT input_valid_d THEN
    channel_fault_d := channel_fault_d + 1;
END_IF;
vote_ok := TwoOfFour(cond_a, cond_b, cond_c, cond_d);
IF cond_a <> cond_b THEN
    diagnosis_count := diagnosis_count + 1;
END_IF;
IF cond_c <> cond_d THEN
    diagnosis_count := diagnosis_count + 1;
END_IF;
IF NOT vote_ok THEN
    diagnosis_count := diagnosis_count + 1;
END_IF;
latch_a_125 := RS_Next(vote_ok, train_a_reset, latch_a_125);
IF latch_a_125 AND (NOT train_a_inhibit) THEN
    mask_a_15 := mask_a_15 + 32;
    trip_a := 0 < 1;
    scram_a := 0 < 1;
    breaker_a := 0 > 1;
    ci_a := 0 < 1;
    alarm_a := 0 < 1;
END_IF;
latch_b_125 := RS_Next(vote_ok, train_b_reset, latch_b_125);
IF latch_b_125 AND (NOT train_b_inhibit) THEN
    mask_b_15 := mask_b_15 + 32;
    trip_b := 0 < 1;
    scram_b := 0 < 1;
    breaker_b := 0 > 1;
    ci_b := 0 < 1;
    alarm_b := 0 < 1;
END_IF;
IF (raw_125_a > 105) AND (NOT cond_a) THEN
    channel_fault_a := channel_fault_a + 1;
END_IF;
IF (raw_125_b > 105) AND (NOT cond_b) THEN
    channel_fault_b := channel_fault_b + 1;
END_IF;
IF (raw_125_c > 105) AND (NOT cond_c) THEN
    channel_fault_c := channel_fault_c + 1;
END_IF;
IF (raw_125_d > 105) AND (NOT cond_d) THEN
    channel_fault_d := channel_fault_d + 1;
END_IF;
IF vote_ok AND train_a_inhibit THEN
    diagnosis_count := diagnosis_count + 1;
END_IF;
IF vote_ok AND train_b_inhibit THEN
    diagnosis_count := diagnosis_count + 1;
END_IF;

cond_a := LimitHigh(raw_126_a, 106);
cond_a := cond_a AND quality_a;
cond_a := cond_a AND (NOT bypass_a);
input_valid_a := InputValid(raw_126_a, 0, 1000);
cond_a := cond_a AND input_valid_a;
IF NOT input_valid_a THEN
    channel_fault_a := channel_fault_a + 1;
END_IF;
cond_b := LimitHigh(raw_126_b, 106);
cond_b := cond_b AND quality_b;
cond_b := cond_b AND (NOT bypass_b);
input_valid_b := InputValid(raw_126_b, 0, 1000);
cond_b := cond_b AND input_valid_b;
IF NOT input_valid_b THEN
    channel_fault_b := channel_fault_b + 1;
END_IF;
cond_c := LimitHigh(raw_126_c, 106);
cond_c := cond_c AND quality_c;
cond_c := cond_c AND (NOT bypass_c);
input_valid_c := InputValid(raw_126_c, 0, 1000);
cond_c := cond_c AND input_valid_c;
IF NOT input_valid_c THEN
    channel_fault_c := channel_fault_c + 1;
END_IF;
cond_d := LimitHigh(raw_126_d, 106);
cond_d := cond_d AND quality_d;
cond_d := cond_d AND (NOT bypass_d);
input_valid_d := InputValid(raw_126_d, 0, 1000);
cond_d := cond_d AND input_valid_d;
IF NOT input_valid_d THEN
    channel_fault_d := channel_fault_d + 1;
END_IF;
vote_ok := TwoOfFour(cond_a, cond_b, cond_c, cond_d);
IF cond_a <> cond_b THEN
    diagnosis_count := diagnosis_count + 1;
END_IF;
IF cond_c <> cond_d THEN
    diagnosis_count := diagnosis_count + 1;
END_IF;
IF NOT vote_ok THEN
    diagnosis_count := diagnosis_count + 1;
END_IF;
latch_a_126 := RS_Next(vote_ok, train_a_reset, latch_a_126);
IF latch_a_126 AND (NOT train_a_inhibit) THEN
    mask_a_15 := mask_a_15 + 64;
    trip_a := 0 < 1;
    scram_a := 0 < 1;
    breaker_a := 0 > 1;
    mfw_a := 0 < 1;
    alarm_a := 0 < 1;
END_IF;
latch_b_126 := RS_Next(vote_ok, train_b_reset, latch_b_126);
IF latch_b_126 AND (NOT train_b_inhibit) THEN
    mask_b_15 := mask_b_15 + 64;
    trip_b := 0 < 1;
    scram_b := 0 < 1;
    breaker_b := 0 > 1;
    mfw_b := 0 < 1;
    alarm_b := 0 < 1;
END_IF;
IF (raw_126_a > 106) AND (NOT cond_a) THEN
    channel_fault_a := channel_fault_a + 1;
END_IF;
IF (raw_126_b > 106) AND (NOT cond_b) THEN
    channel_fault_b := channel_fault_b + 1;
END_IF;
IF (raw_126_c > 106) AND (NOT cond_c) THEN
    channel_fault_c := channel_fault_c + 1;
END_IF;
IF (raw_126_d > 106) AND (NOT cond_d) THEN
    channel_fault_d := channel_fault_d + 1;
END_IF;
IF vote_ok AND train_a_inhibit THEN
    diagnosis_count := diagnosis_count + 1;
END_IF;
IF vote_ok AND train_b_inhibit THEN
    diagnosis_count := diagnosis_count + 1;
END_IF;

cond_a := LimitHigh(raw_127_a, 107);
cond_a := cond_a AND quality_a;
cond_a := cond_a AND (NOT bypass_a);
input_valid_a := InputValid(raw_127_a, 0, 1000);
cond_a := cond_a AND input_valid_a;
IF NOT input_valid_a THEN
    channel_fault_a := channel_fault_a + 1;
END_IF;
cond_b := LimitHigh(raw_127_b, 107);
cond_b := cond_b AND quality_b;
cond_b := cond_b AND (NOT bypass_b);
input_valid_b := InputValid(raw_127_b, 0, 1000);
cond_b := cond_b AND input_valid_b;
IF NOT input_valid_b THEN
    channel_fault_b := channel_fault_b + 1;
END_IF;
cond_c := LimitHigh(raw_127_c, 107);
cond_c := cond_c AND quality_c;
cond_c := cond_c AND (NOT bypass_c);
input_valid_c := InputValid(raw_127_c, 0, 1000);
cond_c := cond_c AND input_valid_c;
IF NOT input_valid_c THEN
    channel_fault_c := channel_fault_c + 1;
END_IF;
cond_d := LimitHigh(raw_127_d, 107);
cond_d := cond_d AND quality_d;
cond_d := cond_d AND (NOT bypass_d);
input_valid_d := InputValid(raw_127_d, 0, 1000);
cond_d := cond_d AND input_valid_d;
IF NOT input_valid_d THEN
    channel_fault_d := channel_fault_d + 1;
END_IF;
vote_ok := TwoOfFour(cond_a, cond_b, cond_c, cond_d);
IF cond_a <> cond_b THEN
    diagnosis_count := diagnosis_count + 1;
END_IF;
IF cond_c <> cond_d THEN
    diagnosis_count := diagnosis_count + 1;
END_IF;
IF NOT vote_ok THEN
    diagnosis_count := diagnosis_count + 1;
END_IF;
latch_a_127 := RS_Next(vote_ok, train_a_reset, latch_a_127);
IF latch_a_127 AND (NOT train_a_inhibit) THEN
    mask_a_15 := mask_a_15 + 128;
    trip_a := 0 < 1;
    scram_a := 0 < 1;
    breaker_a := 0 > 1;
    afw_a := 0 < 1;
    alarm_a := 0 < 1;
END_IF;
latch_b_127 := RS_Next(vote_ok, train_b_reset, latch_b_127);
IF latch_b_127 AND (NOT train_b_inhibit) THEN
    mask_b_15 := mask_b_15 + 128;
    trip_b := 0 < 1;
    scram_b := 0 < 1;
    breaker_b := 0 > 1;
    afw_b := 0 < 1;
    alarm_b := 0 < 1;
END_IF;
IF (raw_127_a > 107) AND (NOT cond_a) THEN
    channel_fault_a := channel_fault_a + 1;
END_IF;
IF (raw_127_b > 107) AND (NOT cond_b) THEN
    channel_fault_b := channel_fault_b + 1;
END_IF;
IF (raw_127_c > 107) AND (NOT cond_c) THEN
    channel_fault_c := channel_fault_c + 1;
END_IF;
IF (raw_127_d > 107) AND (NOT cond_d) THEN
    channel_fault_d := channel_fault_d + 1;
END_IF;
IF vote_ok AND train_a_inhibit THEN
    diagnosis_count := diagnosis_count + 1;
END_IF;
IF vote_ok AND train_b_inhibit THEN
    diagnosis_count := diagnosis_count + 1;
END_IF;

IF trip_a THEN
    trip_counter_a := trip_counter_a + 1;
END_IF;
IF trip_b THEN
    trip_counter_b := trip_counter_b + 1;
END_IF;
IF train_a_reset THEN
    state_a := 0 + 0;
ELSIF trip_a THEN
    state_a := 2 + 0;
ELSIF state_a = 0 THEN
    state_a := 1 + 0;
END_IF;
IF train_b_reset THEN
    state_b := 0 + 0;
ELSIF trip_b THEN
    state_b := 2 + 0;
ELSIF state_b = 0 THEN
    state_b := 1 + 0;
END_IF;

(* ==== FUNCTION_BLOCK 状态输出（用于调试与验证）==== *)
PRINT('FB_DIAG t=', cycle_counter,
      ' pid_pow.U,=', pid_power.U, ' pid_pow.UI,=', pid_power.UI,
      ' pid_tmp.U,=', pid_temp.U, ' pid_tmp.UI,=', pid_temp.UI,
      ' pid_prs.U,=', pid_press.U, ' pid_prs.UI,=', pid_press.UI,
      ' fby_pow.Y,=', fby_power_rate.Y, ' fby_tmp.Y,=', fby_temp_rate.Y,
      ' flt_a.Y,=', filter_fb_a.Y, ' flt_b.Y,=', filter_fb_b.Y,
      ' rs_a.Q,=', rs_prot_a.Q, ' rs_b.Q,=', rs_prot_b.Q,
      ' sr_a.Q,=', sr_reset_a.Q, ' sr_b.Q,=', sr_reset_b.Q,
      '\n');

END_PROGRAM

(* ================================================================
   FUNCTION_BLOCK 定义（v1.5 原生 FB 支持）

   模拟实际核电 RPS 工程中的典型算法块：
     RS_FB      : 置位优先双稳态（保护锁存）
     SR_FB      : 复位优先双稳态（复位控制）
     PID_FB     : 增量式 PID 控制器（功率/温度/压力调节）
     FBY_FB     : 速率限制跟随器（变化率保护）
     FILTER_FB  : 一阶低通滤波器（信号平滑）
   ================================================================ *)

(* ---- RS_FB: 置位优先双稳态（Set-Reset Flip-Flop）---- *)
(* 用于保护通道跳闸锁存，S 与 R 同时为真时输出 1 *)
FUNCTION_BLOCK RS_FB
VAR_INPUT
    S : BOOL;  (* 置位输入：保护条件触发 *)
    R : BOOL;  (* 复位输入：系统复位信号 *)
END_VAR
VAR_OUTPUT
    Q  : BOOL;  (* 正常输出 *)
    QN : BOOL;  (* 反相输出 *)
END_VAR
    Q := S OR (Q AND NOT R);
    QN := NOT Q;
END_FUNCTION_BLOCK

(* ---- SR_FB: 复位优先双稳态（Set-Reset Flip-Flop）---- *)
(* 用于复位控制逻辑，S 与 R 同时为真时输出 0 *)
FUNCTION_BLOCK SR_FB
VAR_INPUT
    S : BOOL;  (* 置位输入 *)
    R : BOOL;  (* 复位输入：优先 *)
END_VAR
VAR_OUTPUT
    Q  : BOOL;
    QN : BOOL;
END_VAR
    Q := (S OR Q) AND NOT R;
    QN := NOT Q;
END_FUNCTION_BLOCK

(* ---- PID_FB: 增量式 PID 控制器 ---- *)
(* 用于反应堆功率、温度、压力调节回路
   特性：
     - 积分项抗饱和（UI 限制在 [UI_LO, UI_HI]）
     - 输出限幅（U 限制在 [LO, HI]）
     - 微分项基于误差变化率（DE = E - E_OLD）
     - VAR_IN_OUT TRACE 用于诊断追踪（直写调用方全局变量）
*)
FUNCTION_BLOCK PID_FB
VAR_INPUT
    E     : DINT;   (* 当前误差 = 设定值 - 测量值 *)
    KP    : DINT;   (* 比例增益 *)
    KD    : DINT;   (* 微分增益 *)
    UI_LO : DINT;   (* 积分项下限 *)
    UI_HI : DINT;   (* 积分项上限 *)
    LO    : DINT;   (* 输出下限 *)
    HI    : DINT;   (* 输出上限 *)
END_VAR
VAR_OUTPUT
    U   : DINT;   (* 控制输出 *)
    UI  : DINT;   (* 积分项当前值 *)
    ALM : BOOL;   (* 输出饱和报警 *)
END_VAR
VAR_IN_OUT
    TRACE : DINT;   (* 诊断追踪：输出同步写入调用方全局 *)
END_VAR
VAR
    DE    : DINT;   (* 误差变化量 *)
    V     : DINT;   (* 积分项临时值 *)
    E_OLD : DINT;   (* 上周期误差 *)
END_VAR
    DE := E - E_OLD;
    V := UI + E;
    IF V > UI_HI THEN
        V := UI_HI;
    ELSIF V < UI_LO THEN
        V := UI_LO;
    END_IF;
    UI := V;
    U := KP * E + UI + KD * DE;
    IF U > HI THEN
        U := HI;
    ELSIF U < LO THEN
        U := LO;
    END_IF;
    IF U >= HI THEN
        ALM := TRUE;
    ELSE
        ALM := FALSE;
    END_IF;
    TRACE := U;
    E_OLD := E;
END_FUNCTION_BLOCK

(* ---- FBY_FB: 速率限制跟随器（First Order Rate Limiter）---- *)
(* 用于保护信号变化率监测，限制信号每周期最大变化量 *)
FUNCTION_BLOCK FBY_FB
VAR_INPUT
    IN : DINT;   (* 输入信号 *)
    DR : DINT;   (* 最大允许变化率（每周期） *)
END_VAR
VAR_OUTPUT
    Y : DINT;   (* 速率限制后的输出 *)
END_VAR
VAR
    V : DINT;   (* 临时值 *)
END_VAR
    V := IN;
    IF V > Y + DR THEN
        V := Y + DR;
    ELSIF V < Y - DR THEN
        V := Y - DR;
    END_IF;
    Y := V;
END_FUNCTION_BLOCK

(* ---- FILTER_FB: 一阶低通滤波器 ---- *)
(* 用于模拟量输入信号平滑处理
   算法：Y_new = Y_old + (IN - Y_old) / ALPHA
   ALPHA 为滤波系数（越大越平滑）
*)
FUNCTION_BLOCK FILTER_FB
VAR_INPUT
    IN    : DINT;   (* 原始输入信号 *)
    ALPHA : DINT;   (* 滤波系数（建议 2-10） *)
END_VAR
VAR_OUTPUT
    Y     : DINT;   (* 滤波后输出 *)
END_VAR
VAR
    DIFF  : DINT;   (* 差值 *)
END_VAR
    DIFF := IN - Y;
    Y := Y + (DIFF / ALPHA);
END_FUNCTION_BLOCK

FUNCTION LimitHigh : BOOL
VAR_INPUT
    value : DINT;
    high : DINT;
END_VAR
LimitHigh := value > high;
END_FUNCTION

FUNCTION InputValid : BOOL
VAR_INPUT
    value : DINT;
    low : DINT;
    high : DINT;
END_VAR
InputValid := (value >= low) AND (value <= high);
END_FUNCTION

FUNCTION OneOfTwo : BOOL
VAR_INPUT
    input_a : BOOL;
    input_b : BOOL;
END_VAR
OneOfTwo := input_a OR input_b;
END_FUNCTION

FUNCTION TwoOfFour : BOOL
VAR_INPUT
    input_a : BOOL;
    input_b : BOOL;
    input_c : BOOL;
    input_d : BOOL;
END_VAR
TwoOfFour := OneOfTwo(OneOfTwo(OneOfTwo(input_a AND input_b, input_c AND input_d), OneOfTwo(input_a AND input_c, input_b AND input_d)), OneOfTwo(input_a AND input_d, input_b AND input_c));
END_FUNCTION

FUNCTION RS_Next : BOOL
VAR_INPUT
    set_input : BOOL;
    reset_input : BOOL;
    q_previous : BOOL;
END_VAR
RS_Next := (set_input OR q_previous) AND (NOT reset_input);
END_FUNCTION

FUNCTION FilterStep : DINT
VAR_INPUT
    previous : DINT;
    input_value : DINT;
END_VAR
FilterStep := previous + ((input_value - previous) / 2);
END_FUNCTION

(* ---- algo_blocks_lib.st ---- *)
(* ================================================================
   algo_blocks_lib.st — SafeST 算法块库（源码级库文件）

   提供 4 种经典控制算法块，全部实现为无状态 FUNCTION：
     RS      : 置位优先双稳态   Q' = S OR (Q_old AND NOT R)
     SR      : 复位优先双稳态   Q' = (S OR Q_old) AND NOT R
     PID_UI  : 积分项 + 限幅    V = UI + KI*E, clamp [LO,HI]
     PID_OUT : 全量输出 + 限幅  U = KP*E + UI + KD*DE, clamp [LO,HI]
     FBY     : 速率限制(跟随)   Q = IN, clamp [PRE-DR, PRE+DR]

   多实例约定（与 rs_multi_entity.st 相同）：
   - 状态（Q_old / UI / DE / PRE）由调用方持有并作为输入传入，
     返回值由调用方写回自身状态变量 => 同一份代码服务任意多个实例。
   - 跨周期状态必须放 VAR_GLOBAL（VM 每周期清零 PROGRAM 局部变量）。
   - 本文件为库源码：VeriSTC 无 LIBRARY/IMPORT 链接机制，
     使用时由上游预处理器将 FUNCTION 块文本内联进目标 .st，
     参见 algo_blocks_multi_instance.st（已内联的可编译测试用例）。
   ================================================================ *)

(* ---- RS：置位优先（S 与 R 同时为真时输出 1） ---- *)
FUNCTION RS : BOOL
VAR_INPUT
  Q_old : BOOL;
  S : BOOL;
  R : BOOL;
END_VAR
  RS := S OR (Q_old AND NOT R);
END_FUNCTION

(* ---- SR：复位优先（S 与 R 同时为真时输出 0） ---- *)
FUNCTION SR : BOOL
VAR_INPUT
  Q_old : BOOL;
  S : BOOL;
  R : BOOL;
END_VAR
  SR := (S OR Q_old) AND NOT R;
END_FUNCTION

(* ---- PID_UI：积分项累加 + 抗积分饱和限幅 ---- *)
FUNCTION PID_UI : DINT
VAR_INPUT
  E  : DINT;
  UI : DINT;
  KI : DINT;
  LO : DINT;
  HI : DINT;
END_VAR
VAR
  V : DINT;
END_VAR
  V := UI + KI * E;
  IF V > HI THEN
    V := HI;
  ELSIF V < LO THEN
    V := LO;
  END_IF;
  PID_UI := V;
END_FUNCTION

(* ---- PID_OUT：比例+积分+微分合成输出 + 限幅 ---- *)
FUNCTION PID_OUT : DINT
VAR_INPUT
  E   : DINT;
  UI  : DINT;
  DE  : DINT;
  KP  : DINT;
  KD  : DINT;
  LO  : DINT;
  HI  : DINT;
END_VAR
VAR
  U : DINT;
END_VAR
  U := KP * E + UI + KD * DE;
  IF U > HI THEN
    U := HI;
  ELSIF U < LO THEN
    U := LO;
  END_IF;
  PID_OUT := U;
END_FUNCTION

(* ---- FBY：一阶速率限制跟随（首出/后备跟随类） ---- *)
FUNCTION FBY : DINT
VAR_INPUT
  IN  : DINT;
  PRE : DINT;
  DR  : DINT;
END_VAR
VAR
  Q : DINT;
END_VAR
  Q := IN;
  IF Q > PRE + DR THEN
    Q := PRE + DR;
  ELSIF Q < PRE - DR THEN
    Q := PRE - DR;
  END_IF;
  FBY := Q;
END_FUNCTION

(* ---- algo_blocks_fb.st ---- *)
(* ================================================================
   algo_blocks_fb.st
   原生 FUNCTION_BLOCK 版算法块库 + "不同变量调用相同算法功能" e2e

   与 FUNCTION 版（algo_blocks_lib.st / algo_blocks_multi_instance.st）
   同激励、同黄金时间线，可交叉验证两种实现一致。

   演示 FB 全部可用特性（P1 + v1.5）：
     - VAR_INPUT / VAR_OUTPUT（多输出：Q 与 QN、U 与 UI 与 ALM）
     - VAR 实例内持久状态（UI / E_OLD，FB_DATA 跨周期不清零）
     - VAR_IN_OUT 逐引用别名（TRACE：诊断量直写调用方全局）
     - 实例声明分离：rs1/rs2 同一份代码、独立数据段
     - IF/ELSIF/ELSE 控制流、表达式实参、命名实参（:=）
   限制：FB 体内不得声明成员实例（嵌套 FB 不支持，P1 范围外）。
   调用点在外部以 IEC 点号访问 inst.FIELD 读取字段（v1.5.1；编译器内部
   融合为不可书写的派生名 inst#FIELD，外部只能读 VAR_OUTPUT）。

   黄金时间线（数值列与 FUNCTION 版一致，t: rs1 rs2 sr1 sr2 | u1 ui1 |
   u2 ui2 | f1 f2，u 与 tr 恒等因 TRACE 别名）。列标签自 v1.5.1 起写作
   点号形式（rs1.Q / pid1.U / pid1.UI / fby1.Y …）指认"这一列来自哪个
   实例的哪个字段"；golden 文件随之只改标签文本，12 行数值逐列不变：
     t1 : 1 0 0 0 | 170 118 | 140 65  |  20   0
     t2 : 1 0 0 0 | 170 200 | 140 90  |  40   0
     t3 : 1 1 0 0 | 170 200 | 140 90  |  60   0
     t4 : 1 0 0 0 | 170 200 | 140 90  |  80   0
     t5 : 0 0 0 0 | 170 200 | 140 90  | 100  50
     t6 : 0 0 0 1 | 170 200 | 140 90  | 120 100
     t7 : 0 0 0 1 | 170 200 | 140 90  | 140 120
     t8 : 0 0 0 1 | 170 200 | 140 90  | 160 120
     t9 : 0 0 0 0 | 170 200 | 135 90  | 180 120
     t10: 0 0 0 0 | 170 200 | 125 90  | 200 120
     t11: 0 0 0 0 | 170 198 | 115 90  | 220 120
     t12: 0 0 0 0 | 158 184 | 105 90  | 240 120
   ================================================================ *)

(* ---- 实例声明：必须先于 POU 列表；每实例独立 FB_DATA ---- *)
VAR_GLOBAL
  rs1  : RS_FB;
  rs2  : RS_FB;
  sr1  : SR_FB;
  sr2  : SR_FB;
  pid1 : PID_FB;
  pid2 : PID_FB;
  fby1 : FBY_FB;
  fby2 : FBY_FB;
  trace1 : DINT;   (* pid1 的 VAR_IN_OUT 别名目标 *)
  trace2 : DINT;   (* pid2 的 VAR_IN_OUT 别名目标 *)
END_VAR

(* ---- RS：置位优先双稳态；Q 为实例持久状态 ---- *)
FUNCTION_BLOCK RS_FB
VAR_INPUT
  S : BOOL;
  R : BOOL;
END_VAR
VAR_OUTPUT
  Q  : BOOL;
  QN : BOOL;
END_VAR
  Q := S OR (Q AND NOT R);
  QN := NOT Q;
END_FUNCTION_BLOCK

(* ---- SR：复位优先双稳态 ---- *)
FUNCTION_BLOCK SR_FB
VAR_INPUT
  S : BOOL;
  R : BOOL;
END_VAR
VAR_OUTPUT
  Q  : BOOL;
  QN : BOOL;
END_VAR
  Q := (S OR Q) AND NOT R;
  QN := NOT Q;
END_FUNCTION_BLOCK

(* ---- PID：定点 PID，实例内持久 UI/E_OLD，KI 固定为 1；
       TRACE 为 VAR_IN_OUT 诊断别名，输出 U 同步写入调用方全局 ---- *)
FUNCTION_BLOCK PID_FB
VAR_INPUT
  E     : DINT;
  KP    : DINT;
  KD    : DINT;
  UI_LO : DINT;
  UI_HI : DINT;
  LO    : DINT;
  HI    : DINT;
END_VAR
VAR_OUTPUT
  U   : DINT;
  UI  : DINT;
  ALM : BOOL;
END_VAR
VAR_IN_OUT
  TRACE : DINT;
END_VAR
VAR
  DE    : DINT;
  V     : DINT;
  E_OLD : DINT;
END_VAR
  DE := E - E_OLD;
  V := UI + E;
  IF V > UI_HI THEN
    V := UI_HI;
  ELSIF V < UI_LO THEN
    V := UI_LO;
  END_IF;
  UI := V;
  U := KP * E + UI + KD * DE;
  IF U > HI THEN
    U := HI;
  ELSIF U < LO THEN
    U := LO;
  END_IF;
  IF U >= HI THEN
    ALM := TRUE;
  ELSE
    ALM := FALSE;
  END_IF;
  TRACE := U;
  E_OLD := E;
END_FUNCTION_BLOCK

(* ---- FBY：速率限制跟随；Y 为实例持久输出 ---- *)
FUNCTION_BLOCK FBY_FB
VAR_INPUT
  IN : DINT;
  DR : DINT;
END_VAR
VAR_OUTPUT
  Y : DINT;
END_VAR
VAR
  V : DINT;
END_VAR
  V := IN;
  IF V > Y + DR THEN
    V := Y + DR;
  ELSIF V < Y - DR THEN
    V := Y - DR;
  END_IF;
  Y := V;
END_FUNCTION_BLOCK

PROGRAM MAIN
VAR
  tick : DINT;
  in2  : DINT;
END_VAR
  tick := CycleCounter();

  (* 与 FUNCTION 版完全相同的激励时序 *)
  rs1(S := (tick = 1), R := (tick = 5));
  rs2(S := (tick = 3), R := (tick = 4));

  sr1(S := (tick = 2), R := (tick = 2));
  sr2(S := (tick = 6), R := (tick = 9));

  (* 同一份 PID 代码，两套增益/限值、两套独立状态与别名目标 *)
  pid1(E := 130 - tick * 12, KP := 1, KD := 1,
       UI_LO := 0, UI_HI := 200, LO := 0, HI := 170,
       TRACE := trace1);
  pid2(E := 70 - tick * 5, KP := 2, KD := 1,
       UI_LO := 0, UI_HI := 90, LO := 0, HI := 140,
       TRACE := trace2);

  fby1(IN := tick * 30, DR := 20);
  IF tick > 4 THEN
    in2 := 120;
  ELSE
    in2 := 0;
  END_IF;
  fby2(IN := in2, DR := 50);

  PRINT('FB t=', tick, ' rs1.Q,=', rs1.Q, ' rs2.Q,=', rs2.Q,
        ' sr1.Q,=', sr1.Q, ' sr2.Q,=', sr2.Q,
        ' pid1.U,=', pid1.U, ' pid1.UI,=', pid1.UI,
        ' pid2.U,=', pid2.U, ' pid2.UI,=', pid2.UI,
        ' fby1.Y,=', fby1.Y, ' fby2.Y,=', fby2.Y,
        ' trace1,=', trace1, ' trace2,=', trace2, '\n');
END_PROGRAM

(* ---- native_fb_in_out.st ---- *)
(* ================================================================
   native_fb_in_out.st  --  VAR_IN_OUT 逐引用别名 e2e

   验证 v1.5 IN_OUT 语义：端口不是副本，而是调用方存储的别名。
     - 逻辑一份（ACCUM 定义），实例数据分离（a1/a2 各自持有 LAST）
     - VAR_IN_OUT ACC 编译为"指向调用方全局的地址"形参，体内读写走
       I32_LOAD_PTR / I32_STORE_PTR，故两个实例共享同一个 shared
     - 同一周期内双向可见：调用方写 shared → 被调读得到；被调写
       ACC → 调用方立即读到

   每周期 t（tick = CycleCounter()）：
     shared := t                 调用方写入别名目标
     a1(K := 10)  : LAST := t,       shared := t + 10
     a2(K := 100) : LAST := t + 10,  shared := t + 110
   ⇒ PRINT 输出 (tick, shared, a1.LAST, a2.LAST)
        t=1 → 1, 111, 1, 11     t=3 → 3, 113, 3, 13
   LAST 互不相同 ⇒ 实例数据仍分离；shared 单点累加 ⇒ 端口是别名。
   ================================================================ *)

(* 实例声明必须先于 POU 列表（顶层文法：VAR_GLOBAL → POU*）*)
VAR_GLOBAL
  shared : DINT;
  a1 : ACCUM;
  a2 : ACCUM;
END_VAR

FUNCTION_BLOCK ACCUM
VAR_INPUT
  K : DINT;
END_VAR
VAR_OUTPUT
  LAST : DINT;
END_VAR
VAR_IN_OUT
  ACC : DINT;
END_VAR
  LAST := ACC;
  ACC := ACC + K;
END_FUNCTION_BLOCK

PROGRAM MAIN
VAR
  tick : DINT;
END_VAR
  tick := CycleCounter();
  shared := tick;
  a1(ACC := shared, K := 10);
  a2(ACC := shared, K := 100);
  PRINT('tick', tick, shared, a1.LAST, a2.LAST);
END_PROGRAM

(* ---- native_fb_multi_instance.st ---- *)
(* ================================================================
   native_fb_multi_instance.st  --  原生 FUNCTION_BLOCK 多实体 e2e

   验证 P1 目标：库逻辑一份（FB 定义），实例数据分离（每实例
   独立 self 相对上下文），无需前端文本预处理器展开。

   语义（RS，S 置位优先于 R 复位）： Q := S OR (Q AND NOT R)
     - 逻辑体只在 FUNCTION_BLOCK RS_V1 出现一份
     - rs1 / rs2 为两个实例，各自持有独立的 Q 上下文
     - MAIN 只见调用与实例输出读取，不复制算法体

   tick = CycleCounter(): 1,2,3,...
   rs1: S=(tick=2) R=(tick=6)  -> Q: 0,0,1,1,1,1,0,0
   rs2: S=(tick=4) R=(tick=8)  -> Q: 0,0,0,1,1,1,1,0
   ================================================================ *)

(* 实例声明必须先于 POU 列表（顶层文法：VAR_GLOBAL → POU*）*)
VAR_GLOBAL
  rs1 : RS_FB;
  rs2 : RS_FB;
END_VAR

FUNCTION_BLOCK RS_FB
VAR_INPUT
  S : BOOL;
  R : BOOL;
END_VAR
VAR_OUTPUT
  Q : BOOL;
END_VAR
  Q := S OR (Q AND NOT R);
END_FUNCTION_BLOCK

PROGRAM MAIN
VAR
  tick : DINT;
END_VAR
  tick := CycleCounter();
  rs1(S := (tick = 2), R := (tick = 6));
  rs2(S := (tick = 4), R := (tick = 8));
  PRINT('tick', tick, rs1.Q, rs2.Q);
END_PROGRAM

(* ---- qualified_access_field.st ---- *)
(* ================================================================
   qualified_access_field.st -- IEC 点号访问 + 派生名不可书写 e2e

   验证 v1.5.1 两项改动在同一程序里共存且互不干扰：
     1) inst.field（此处 l1.Q）由 parser 就地融合为内部派生名 l1#Q，
        与 expand_instances 生成的扁平全局逐字一致 ⇒ 调用方可以按
        IEC 写法只读实例输出，无需再手写 a1_Q 这类扁平名；
     2) 分隔符 '#' 不在标识符文法（字母 (字母|数字|_)*）内 ⇒ 派生名
        不可书写：用户既写不出 l1#Q（词法即报错），也不能拿它冒充
        自己声明的名字。同名风格的扁平全局 l1_Q 因此只是一个普通变量。

   语义：
     l1 : LATCH，体内 C := C + 1（私有状态）、Q := K + 1（输出）
     tick = CycleCounter(): 1,2,3,...
     l1(K := tick)          ⇒ l1.Q  = tick + 1
     l1_Q := 100 * tick     ⇒ 用户全局，与实例字段无关
   ⇒ PRINT 输出 (tick, l1_Q, l1.Q)
        t=1 → 1, 100, 2    t=2 → 2, 200, 3    t=4 → 4, 400, 5
   两条轨迹同步而不合并 ⇒ 名字空间已分离。
   反向用例（写 l1.Q / 读 l1.C）见 negative/qualified_*.st。
   ================================================================ *)

VAR_GLOBAL
  l1 : LATCH;
  l1_Q : DINT;
END_VAR

FUNCTION_BLOCK LATCH
VAR_INPUT
  K : DINT;
END_VAR
VAR_OUTPUT
  Q : DINT;
END_VAR
VAR
  C : DINT;
END_VAR
  C := C + 1;
  Q := K + 1;
END_FUNCTION_BLOCK

PROGRAM MAIN
VAR
  tick : DINT;
END_VAR
  tick := CycleCounter();
  l1(K := tick);
  l1_Q := 100 * tick;
  PRINT('tick', tick, l1_Q, l1.Q);
END_PROGRAM

(* ---- sim_closed_loop.st ---- *)
(* ================================================================
   sim_closed_loop.st -- closed-loop demo for the simulation backend

   An integral controller against a first-order-lag plant. Three signals
   cross the I/O boundary:

     pv : AI ch0 -- the controlled quantity, produced by the plant
     mv : AO ch1 -- the manipulated value, written by the controller
     sp : AI ch2 -- the setpoint, a constant source in the plant

   The controller is deliberately written with DINT only (decision D1: the
   REAL chain is not usable yet), so units are integer counts over 0..1000
   and the loop is closed by the simulator, not by ST.

   Anti-windup: the accumulator integrates only while inside its bounds and
   is clamped afterwards, since integrator + saturated actuator otherwise
   winds up and the loop never recovers.

   Golden timeline (12 cycles, period 100 ms, plant gain 1/8), recorded from
   build/bin/sim and diffed by integration/run_sim_e2e.sh. The values shown
   are the ones the channel carried at the start of that cycle:
     cycle  sp   pv   mv
         1 500    0  500
         2 500   62  938
         3 500  171 1000
         4 500  274 1000
         5 500  364 1000
         6 500  443 1000
         7 500  512  988
         8 500  571  917
         9 500  614  803
        10 500  637  666
        11 500  640  526
        12 500  625  401
   The actuator saturates for four cycles, the accumulator stops winding up
   there, and the controlled quantity turns back toward the setpoint on its
   own: a closed loop with no operator and no wall clock.

   `cnt` exists for the watch layer only (G0 deliverable 4): a FUNCTION_BLOCK
   instance whose fields land in the symbol table as derived names
   `cnt#N` / `cnt#ACC`, so integration/run_sim_e2e.sh can prove that watching
   an instance field resolves through section 7 to a live slot. It is called
   once per cycle with STEP := 1 and touches none of the loop signals, which
   is why the timeline above is unchanged by adding it.
   ================================================================ *)

VAR_GLOBAL
  sp    : DINT;
  pv    : DINT;
  mv    : DINT;
  err   : DINT;
  integ : DINT;
  cnt   : COUNTER_FB;
END_VAR
IOMAP
  pv, 0, INPUT, DINT;
  mv, 1, OUTPUT, DINT;
  sp, 2, INPUT, DINT;
END_IOMAP
(* 每周期 +STEP，N 是对外可见的累计值，ACC 是实例内部状态 *)
FUNCTION_BLOCK COUNTER_FB
VAR_INPUT
  STEP : DINT;
END_VAR
VAR_OUTPUT
  N : DINT;
END_VAR
VAR
  ACC : DINT;
END_VAR
  ACC := ACC + STEP;
  N := ACC;
END_FUNCTION_BLOCK
PROGRAM MAIN
  err := sp - pv;
  cnt(STEP := 1);

  IF (err > 0) AND (integ < 1000) THEN
    integ := integ + err;
  END_IF;

  IF (err < 0) AND (integ > 0) THEN
    integ := integ + err;
  END_IF;

  IF integ > 1000 THEN
    integ := 1000;
  END_IF;

  IF integ < 0 THEN
    integ := 0;
  END_IF;

  mv := integ;
END_PROGRAM

(* ---- algo_blocks_multi_instance.st ---- *)
(* ================================================================
   algo_blocks_multi_instance.st
   测试用例：不同的变量调用相同的算法功能（多实例复用）

   内联库：tests/st-examples/algo_blocks_lib.st
   （VeriSTC 无库链接机制，库文本由上游预处理器内联，此处手工内联）

   每个算法块均有 2 个实例，实例之间变量完全独立：
     RS(q1)/RS(q2)   SR(q1)/SR(q2)
     PID(e1,ui1,de1,u1) / PID(e2,ui2,de2,u2)
     FBY(in->f1) / FBY(in->f2)
   跨周期状态全部放 VAR_GLOBAL 并由调用方写回。

   12 周期金标准（t: rs1 rs2 sr1 sr2 | u1 ui1 | u2 ui2 | f1 f2）
     t1 : 1 0 0 0 | 170 118 | 140 65  |  20   0
     t2 : 1 0 0 0 | 170 200 | 140 90  |  40   0
     t3 : 1 1 0 0 | 170 200 | 140 90  |  60   0
     t4 : 1 0 0 0 | 170 200 | 140 90  |  80   0
     t5 : 0 0 0 0 | 170 200 | 140 90  | 100  50
     t6 : 0 0 0 1 | 170 200 | 140 90  | 120 100
     t7 : 0 0 0 1 | 170 200 | 140 90  | 140 120
     t8 : 0 0 0 1 | 170 200 | 140 90  | 160 120
     t9 : 0 0 0 0 | 170 200 | 135 90  | 180 120
     t10: 0 0 0 0 | 170 200 | 125 90  | 200 120
     t11: 0 0 0 0 | 170 198 | 115 90  | 220 120
     t12: 0 0 0 0 | 158 184 | 105 90  | 240 120
   ================================================================ *)

VAR_GLOBAL
  rs1_q  : BOOL;
  rs2_q  : BOOL;
  sr1_q  : BOOL;
  sr2_q  : BOOL;
  pid1_ui   : DINT;
  pid1_eold : DINT;
  pid2_ui   : DINT;
  pid2_eold : DINT;
  fby1_out : DINT;
  fby2_out : DINT;
END_VAR

(* ---------------- 库：algo_blocks_lib.st 内联开始 ---------------- *)

FUNCTION RS : BOOL
VAR_INPUT
  Q_old : BOOL;
  S : BOOL;
  R : BOOL;
END_VAR
  RS := S OR (Q_old AND NOT R);
END_FUNCTION

FUNCTION SR : BOOL
VAR_INPUT
  Q_old : BOOL;
  S : BOOL;
  R : BOOL;
END_VAR
  SR := (S OR Q_old) AND NOT R;
END_FUNCTION

FUNCTION PID_UI : DINT
VAR_INPUT
  E  : DINT;
  UI : DINT;
  KI : DINT;
  LO : DINT;
  HI : DINT;
END_VAR
VAR
  V : DINT;
END_VAR
  V := UI + KI * E;
  IF V > HI THEN
    V := HI;
  ELSIF V < LO THEN
    V := LO;
  END_IF;
  PID_UI := V;
END_FUNCTION

FUNCTION PID_OUT : DINT
VAR_INPUT
  E   : DINT;
  UI  : DINT;
  DE  : DINT;
  KP  : DINT;
  KD  : DINT;
  LO  : DINT;
  HI  : DINT;
END_VAR
VAR
  U : DINT;
END_VAR
  U := KP * E + UI + KD * DE;
  IF U > HI THEN
    U := HI;
  ELSIF U < LO THEN
    U := LO;
  END_IF;
  PID_OUT := U;
END_FUNCTION

FUNCTION FBY : DINT
VAR_INPUT
  IN  : DINT;
  PRE : DINT;
  DR  : DINT;
END_VAR
VAR
  Q : DINT;
END_VAR
  Q := IN;
  IF Q > PRE + DR THEN
    Q := PRE + DR;
  ELSIF Q < PRE - DR THEN
    Q := PRE - DR;
  END_IF;
  FBY := Q;
END_FUNCTION

(* ---------------- 库内联结束 ---------------- *)

PROGRAM MAIN
VAR
  tick  : DINT;
  rs1_s : BOOL;
  rs1_r : BOOL;
  rs2_s : BOOL;
  rs2_r : BOOL;
  sr1_s : BOOL;
  sr1_r : BOOL;
  sr2_s : BOOL;
  sr2_r : BOOL;
  e1  : DINT;
  de1 : DINT;
  u1  : DINT;
  e2  : DINT;
  de2 : DINT;
  u2  : DINT;
  in1 : DINT;
  in2 : DINT;
  fby1_q : DINT;
  fby2_q : DINT;
END_VAR
  tick := CycleCounter();

  (* ---- 激励 ---- *)
  rs1_s := tick = 1;
  rs1_r := tick = 5;
  rs2_s := tick = 3;
  rs2_r := tick = 4;
  sr1_s := tick = 2;
  sr1_r := tick = 2;
  sr2_s := tick = 6;
  sr2_r := tick = 9;

  (* ---- RS：同一功能，两套变量 ---- *)
  rs1_q := RS(rs1_q, rs1_s, rs1_r);
  rs2_q := RS(rs2_q, rs2_s, rs2_r);

  (* ---- SR：同一功能，另两套变量 ---- *)
  sr1_q := SR(sr1_q, sr1_s, sr1_r);
  sr2_q := SR(sr2_q, sr2_s, sr2_r);

  (* ---- PID 实例 1：e1 = 130 - 12t, Kp=Ki=Kd=1, UI限[0,200], U限[0,170] ---- *)
  e1  := 130 - tick * 12;
  de1 := e1 - pid1_eold;
  pid1_ui := PID_UI(e1, pid1_ui, 1, 0, 200);
  u1  := PID_OUT(e1, pid1_ui, de1, 1, 1, 0, 170);
  pid1_eold := e1;

  (* ---- PID 实例 2：e2 = 70 - 5t, Kp=2,Kd=1, UI限[0,90], U限[0,140] ---- *)
  e2  := 70 - tick * 5;
  de2 := e2 - pid2_eold;
  pid2_ui := PID_UI(e2, pid2_ui, 1, 0, 90);
  u2  := PID_OUT(e2, pid2_ui, de2, 2, 1, 0, 140);
  pid2_eold := e2;

  (* ---- FBY 实例 1：in1 = 30t 斜坡, 速率限 20 ---- *)
  in1 := tick * 30;
  fby1_q := FBY(in1, fby1_out, 20);
  fby1_out := fby1_q;

  (* ---- FBY 实例 2：t<=4 时 in2=0，之后跳变 120, 速率限 50 ---- *)
  IF tick > 4 THEN
    in2 := 120;
  ELSE
    in2 := 0;
  END_IF;
  fby2_q := FBY(in2, fby2_out, 50);
  fby2_out := fby2_q;

  PRINT('ALG t=', tick, ' rs1=', rs1_q, ' rs2=', rs2_q,
        ' sr1=', sr1_q, ' sr2=', sr2_q,
        ' u1=', u1, ' ui1=', pid1_ui,
        ' u2=', u2, ' ui2=', pid2_ui,
        ' f1=', fby1_out, ' f2=', fby2_out, '\n');
END_PROGRAM

(* ---- core_assign.st ---- *)
PROGRAM P
VAR
    x : DINT;
    counter : DINT;
END_VAR
counter := CycleCounter();
x := 42 + 0;
PRINT('counter=', counter, ' x=', x, '\n');
END_PROGRAM

(* ---- function_control_flow.st ---- *)
(* Full stateless FUNCTION support:
   - local variables
   - IF/ELSIF/ELSE control flow
   - nested FUNCTION calls
   - real CALL/RETURN code generation *)

FUNCTION AddOne : DINT
VAR_INPUT
  x : DINT;
END_VAR
  AddOne := x + 1;
END_FUNCTION

FUNCTION Clamp : DINT
VAR_INPUT
  x  : DINT;
  lo : DINT;
  hi : DINT;
END_VAR
VAR
  r : DINT;
END_VAR
  IF x < lo THEN
    r := lo;
  ELSIF x > hi THEN
    r := hi;
  ELSE
    r := x;
  END_IF;
  Clamp := r;
END_FUNCTION

PROGRAM MAIN
VAR
  tick : DINT;
  y    : DINT;
END_VAR
  tick := CycleCounter();
  y := Clamp(AddOne(tick), 2, 5);
  PRINT('tick=', tick, ' y=', y, '\n');
END_PROGRAM

(* ---- function_impure.st ---- *)
(* Negative test: FUNCTION must remain stateless.
   It may not assign to VAR_INPUT or VAR_GLOBAL. *)

VAR_GLOBAL
  g : DINT;
END_VAR

FUNCTION Bad : DINT
VAR_INPUT
  x : DINT;
END_VAR
  x := 1;
  g := 2;
  Bad := x;
END_FUNCTION

PROGRAM MAIN
VAR
  y : DINT;
END_VAR
  y := Bad(0);
  PRINT('y=', y, '\n');
END_PROGRAM

(* ---- function_local_initializer.st ---- *)
(* Positive test: FUNCTION local initializers are lowered to entry assignments.
   Each call re-initializes r before executing the body. *)

FUNCTION Next : DINT
VAR_INPUT
  x : DINT;
END_VAR
VAR
  r : DINT := 10;
END_VAR
  r := r + x;
  Next := r;
END_FUNCTION

PROGRAM MAIN
VAR
  y : DINT;
END_VAR
  y := Next(1);
  PRINT('y=', y, '\n');
END_PROGRAM

(* ---- function_loop.st ---- *)
(* Positive test: constant-bound FOR is allowed inside a stateless FUNCTION.
   WHILE/REPEAT remain rejected until loop-variant analysis is complete. *)

FUNCTION SumTo : DINT
VAR_INPUT
  n : DINT;
END_VAR
VAR
  i : INT;
  s : DINT;
END_VAR
  FOR i := 0 TO 10 DO
    s := s + 1;
  END_FOR;
  SumTo := s;
END_FUNCTION

PROGRAM MAIN
VAR
  y : DINT;
END_VAR
  y := SumTo(3);
  PRINT('y=', y, '\n');
END_PROGRAM

(* ---- function_recursive.st ---- *)
(* Negative test: direct recursion is rejected before code generation. *)

FUNCTION Fact : DINT
VAR_INPUT
  n : DINT;
END_VAR
  Fact := n * Fact(n - 1);
END_FUNCTION

PROGRAM MAIN
VAR
  y : DINT;
END_VAR
  y := Fact(3);
  PRINT('y=', y, '\n');
END_PROGRAM

(* ---- function_while.st ---- *)
(* Negative test: WHILE is not yet allowed inside FUNCTION bodies.
   It requires loop-variant analysis in a call frame and additional proofs. *)

FUNCTION WaitPositive : DINT
VAR_INPUT
  n : DINT;
END_VAR
VAR
  y : DINT;
END_VAR
  WHILE y < n DO
    y := y + 1;
  END_WHILE;
  WaitPositive := y;
END_FUNCTION

PROGRAM MAIN
VAR
  y : DINT;
END_VAR
  y := WaitPositive(3);
  PRINT('y=', y, '\n');
END_PROGRAM

(* ---- io_cal.st ---- *)
(* IOMAP smoke: two mapped channels, one input and one output.
   The IOMAP block is the only place a channel number and direction are
   declared; scale/bias are emitted by the compiler as identity (1.0 / 0.0)
   and the loader must read them from the file instead of hardcoding them. *)
VAR_GLOBAL
    ai0 : DINT;
    ao0 : DINT;
END_VAR
IOMAP
    ai0, 0, INPUT, DINT;
    ao0, 1, OUTPUT, DINT;
END_IOMAP
PROGRAM P
    ao0 := ai0 + 1;
END_PROGRAM

(* ---- nuclear_rps_channel.st ---- *)
(* ================================================================
   nuclear_rps_channel.st — 单组 RPS 4 通道保护 + 跳闸母线 + ESFAS 顺序器

   定位（与 feature-probes/ 分工）：探针覆盖单构造，本文件覆盖
   "状态密集 + 核电保护语义"，全部构造限于当前实编译管线
   （global_codegen I32 后端）可正确执行的子集：
     CASE 多分支(值/范围/ELSE) · IF/ELSIF · FOR(INT 环变量) ·
     WHILE 定点缩放 · MOD/除法 · 布尔代数(AND/OR/XOR/NOT) ·
     FUNCTION 多实参内联复用 · VAR_GLOBAL 跨周期锁存 ·
     CycleCounter 驱动场景激励 · PRINT 可观测量

   被保护对象：核岛 RPS 保护机柜（4 通道 A/B/C/D，中子功率量程，
   整定 1100/堆量程单位，迟滞复位 1000）。跳闸母线 2oo4 表决，
   故障/旁路通道从表决中剔除。ESFAS 顺序器按周期间隔分级：
   SI 信号 → 高压注泵 → 停堆卸压。

   场景时间线（tick = CycleCounter，运行 38 周期）：
     t=11..21  A 通道超量程(1160)
     t=13..23  B 通道超量程(1160)
     t=13..    D 通道持续超量程(1160)
     t=5..8    C 传感器故障(sf_c)  t>=9 C 维护旁路(byp_c)
     t=14/16   A/B/D 滤波均值越限 → 触发延时 3 周期(TON 仿真)
     t=17      A 跳闸  t=19 B/D 跳闸 → 2oo4 满足 → 母线 A 跳
               (上升沿 trip_count_a=1, 顺序器启动)
     t=24 SI, t=28 HPI …  t=30 全局 RESET：闭锁清除、顺序器复位
     t=33      D 重新跳闸，但仅剩 1/4 → 母线保持释放（验证复位后
               表决抑制路径）
   ================================================================ *)

(* ---------------- 跨周期状态（VM 持久 MEM 段） ---------------- *)

VAR_GLOBAL
  (* 通道状态机: 0=NORMAL 2=TRIP_PENDING 3=TRIPPED 4=BYPASSED 5=FAULT *)
  st_a : DINT;
  st_b : DINT;
  st_c : DINT;
  st_d : DINT;
  (* 跳闸延时计时器 (TON 仿真, 单位=扫描周期) *)
  dt_a : DINT;
  dt_b : DINT;
  dt_c : DINT;
  dt_d : DINT;
  (* 4 抽头滑动平均环 × 4 通道 = 16 个状态字 *)
  f0_a : DINT;
  f1_a : DINT;
  f2_a : DINT;
  f3_a : DINT;
  f0_b : DINT;
  f1_b : DINT;
  f2_b : DINT;
  f3_b : DINT;
  f0_c : DINT;
  f1_c : DINT;
  f2_c : DINT;
  f3_c : DINT;
  f0_d : DINT;
  f1_d : DINT;
  f2_d : DINT;
  f3_d : DINT;
  (* 滤波输出 *)
  avg_a : DINT;
  avg_b : DINT;
  avg_c : DINT;
  avg_d : DINT;
  (* 跳闸闭锁 *)
  trip_a : BOOL;
  trip_b : BOOL;
  trip_c : BOOL;
  trip_d : BOOL;
  (* 跳闸母线 + 边沿检测 + 计数器 *)
  trainA_trip : BOOL;
  prevA : BOOL;
  trip_count_a : DINT;
  (* ESFAS 顺序器: 0=IDLE 1=SI延时 2=HPI延时 3=卸压延时 4=完成 *)
  seq_state : DINT;
  seq_timer : DINT;
  si_a : BOOL;
  hpi_a : BOOL;
  ld_a : BOOL;
  (* 报警字 *)
  alarm_word : DINT;
END_VAR

(* ---------------- 库函数（内联展开，多实体复用） ---------------- *)

(* 4 点滑动平均（定点） *)
FUNCTION MA4 : DINT
VAR_INPUT
  x0 : DINT;
  x1 : DINT;
  x2 : DINT;
  x3 : DINT;
END_VAR
  MA4 := (x0 + x1 + x2 + x3) / 4;
END_FUNCTION

(* 2oo3 表决：三输入中至少两个为真 *)
FUNCTION Vote23 : BOOL
VAR_INPUT
  a : BOOL;
  b : BOOL;
  c : BOOL;
END_VAR
  Vote23 := (a AND b) OR (a AND c) OR (b AND c);
END_FUNCTION

(* 通道有效跳闸输出：故障或旁路时强制剔除 *)
FUNCTION ChValid : BOOL
VAR_INPUT
  q : BOOL;
  fault : BOOL;
  bypass : BOOL;
END_VAR
  ChValid := q AND (NOT fault) AND (NOT bypass);
END_FUNCTION

(* ---------------- 主程序 ---------------- *)

PROGRAM MAIN
VAR
  tick : DINT;
  (* 输入层临时量 *)
  raw_a : DINT;
  raw_b : DINT;
  raw_c : DINT;
  raw_d : DINT;
  byp_c : BOOL;
  sf_c : BOOL;
  rst : BOOL;
  (* 表决有效输出 *)
  va : BOOL;
  vb : BOOL;
  vc : BOOL;
  vd : BOOL;
  vote : BOOL;
  (* 报警字打包 / 位重编码 (FOR) *)
  fa : DINT;
  bitv : DINT;
  pow : DINT;
  j : INT;
  (* 定点百分比缩放 (WHILE) *)
  n : DINT;
  pct_a : DINT;
END_VAR
  tick := CycleCounter();

  (* ---- 1. 场景激励（确定性，tick 驱动） ---- *)
  raw_c := 880;
  raw_a := 880;
  IF (tick >= 11) AND (tick <= 21) THEN
    raw_a := 1160;
  END_IF;
  raw_b := 880;
  IF (tick >= 13) AND (tick <= 23) THEN
    raw_b := 1160;
  END_IF;
  raw_d := 880;
  IF tick >= 13 THEN
    raw_d := 1160;
  END_IF;
  sf_c := (tick >= 5) AND (tick <= 8);
  byp_c := tick >= 9;
  rst := tick = 30;

  (* ---- 2. 滑动平均环更新（右旋 + 新样本入 f0） ---- *)
  f3_a := f2_a;
  f2_a := f1_a;
  f1_a := f0_a;
  f0_a := raw_a;
  avg_a := MA4(f0_a, f1_a, f2_a, f3_a);

  f3_b := f2_b;
  f2_b := f1_b;
  f1_b := f0_b;
  f0_b := raw_b;
  avg_b := MA4(f0_b, f1_b, f2_b, f3_b);

  f3_c := f2_c;
  f2_c := f1_c;
  f1_c := f0_c;
  f0_c := raw_c;
  avg_c := MA4(f0_c, f1_c, f2_c, f3_c);

  f3_d := f2_d;
  f2_d := f1_d;
  f1_d := f0_d;
  f0_d := raw_d;
  avg_d := MA4(f0_d, f1_d, f2_d, f3_d);

  (* ---- 3. RESET：清除所有闭锁与顺序器 ---- *)
  IF rst THEN
    st_a := 0;  st_b := 0;  st_d := 0;
    dt_a := 0;  dt_b := 0;  dt_d := 0;
    trip_a := FALSE;  trip_b := FALSE;  trip_d := FALSE;
    trainA_trip := FALSE;
    seq_state := 0;  seq_timer := 0;
    si_a := FALSE;  hpi_a := FALSE;  ld_a := FALSE;
  END_IF;

  (* ---- 4. C 通道维护状态直通（旁路优先于故障） ---- *)
  IF byp_c THEN
    st_c := 4;
  ELSIF sf_c THEN
    st_c := 5;
  ELSE
    st_c := 0;
  END_IF;

  (* ---- 5. 每通道跳闸状态机（多分支 CASE） ----
     NORMAL → 均值越限 → TRIP_PENDING(延时 3 周期) → TRIPPED；
     PENDING 中均值回落则撤回 NORMAL（延时取消）。 *)
  CASE st_a OF
    0:
      IF avg_a > 1100 THEN
        st_a := 2;
        dt_a := 3;
      END_IF;
    2:
      dt_a := dt_a - 1;
      IF dt_a <= 0 THEN
        st_a := 3;
        trip_a := TRUE;
      ELSE
        IF avg_a <= 1000 THEN
          st_a := 0;
        END_IF;
      END_IF;
    3:
      trip_a := TRUE;
    4:
      trip_a := FALSE;
    5:
      trip_a := FALSE;
  END_CASE;

  CASE st_b OF
    0:
      IF avg_b > 1100 THEN
        st_b := 2;
        dt_b := 3;
      END_IF;
    2:
      dt_b := dt_b - 1;
      IF dt_b <= 0 THEN
        st_b := 3;
        trip_b := TRUE;
      ELSE
        IF avg_b <= 1000 THEN
          st_b := 0;
        END_IF;
      END_IF;
    3:
      trip_b := TRUE;
    4:
      trip_b := FALSE;
    5:
      trip_b := FALSE;
  END_CASE;

  CASE st_c OF
    0:
      IF avg_c > 1100 THEN
        st_c := 2;
        dt_c := 3;
      END_IF;
    2:
      dt_c := dt_c - 1;
      IF dt_c <= 0 THEN
        st_c := 3;
        trip_c := TRUE;
      ELSE
        IF avg_c <= 1000 THEN
          st_c := 0;
        END_IF;
      END_IF;
    3:
      trip_c := TRUE;
    4:
      trip_c := FALSE;
    5:
      trip_c := FALSE;
  END_CASE;

  CASE st_d OF
    0:
      IF avg_d > 1100 THEN
        st_d := 2;
        dt_d := 3;
      END_IF;
    2:
      dt_d := dt_d - 1;
      IF dt_d <= 0 THEN
        st_d := 3;
        trip_d := TRUE;
      ELSE
        IF avg_d <= 1000 THEN
          st_d := 0;
        END_IF;
      END_IF;
    3:
      trip_d := TRUE;
    4:
      trip_d := FALSE;
    5:
      trip_d := FALSE;
  END_CASE;

  (* ---- 6. 2oo4 表决（剔除故障/旁路通道） + 母线自保持 + 上升沿 ---- *)
  va := ChValid(trip_a, FALSE, FALSE);
  vb := ChValid(trip_b, FALSE, FALSE);
  vc := ChValid(trip_c, sf_c, byp_c);
  vd := ChValid(trip_d, FALSE, FALSE);
  vote := Vote23(va, vb, vd);
  trainA_trip := trainA_trip OR vote;
  IF trainA_trip AND (NOT prevA) THEN
    trip_count_a := trip_count_a + 1;
    IF seq_state = 0 THEN
      seq_state := 1;
      seq_timer := 5;
    END_IF;
  END_IF;
  prevA := trainA_trip;

  (* ---- 7. ESFAS 顺序器（周期分级延时） ---- *)
  IF seq_state = 1 THEN
    seq_timer := seq_timer - 1;
    IF seq_timer <= 0 THEN
      si_a := TRUE;
      seq_state := 2;
      seq_timer := 4;
    END_IF;
  ELSIF seq_state = 2 THEN
    seq_timer := seq_timer - 1;
    IF seq_timer <= 0 THEN
      hpi_a := TRUE;
      seq_state := 3;
      seq_timer := 4;
    END_IF;
  ELSIF seq_state = 3 THEN
    seq_timer := seq_timer - 1;
    IF seq_timer <= 0 THEN
      ld_a := TRUE;
      seq_state := 4;
    END_IF;
  END_IF;

  (* ---- 8. 报警字: bit3=A跳 bit2=B跳 bit1=C故障/旁路 bit0=D跳；
         FOR 环做位域重编码（/·MOD 取位后原样重组，恒等即通过） ---- *)
  fa := 0;
  IF va THEN
    fa := fa + 8;
  END_IF;
  IF vb THEN
    fa := fa + 4;
  END_IF;
  IF sf_c OR byp_c THEN
    fa := fa + 2;
  END_IF;
  IF vd THEN
    fa := fa + 1;
  END_IF;
  alarm_word := 0;
  pow := 1;
  FOR j := 0 TO 3 DO
    bitv := (fa / pow) MOD 2;
    alarm_word := alarm_word + bitv * pow;
    pow := pow * 2;
  END_FOR;

  (* ---- 9. A 通道量程百分比：无浮点定点缩放（WHILE 收敛环） ---- *)
  n := raw_a;
  pct_a := 0;
  WHILE n >= 12 DO
    n := n - 12;
    pct_a := pct_a + 1;
  END_WHILE;

  (* ---- 10. 可观测量 ---- *)
  PRINT('CHAN t=', tick, ' av=', avg_a, ',', avg_b, ',', avg_c, ',', avg_d,
        ' st=', st_a, ',', st_b, ',', st_c, ',', st_d,
        ' v=', va, ',', vb, ',', vc, ',', vd,
        ' bus=', trainA_trip, ' cnt=', trip_count_a,
        ' seq=', seq_state, ',', si_a, ',', hpi_a, ',', ld_a,
        ' aw=', alarm_word, ' pct=', pct_a, '\n');
END_PROGRAM

(* ---- rs_multi_entity.st ---- *)
(* ================================================================
   rs_multi_entity.st
   Multi-entity pattern: ONE function entity (RS bistable) called
   multiple times, each call passing the caller's own variables
   plus its previous state; the single return value is the new
   state, written back by the caller.

     q1 := RS(q1, s1, r1);   (* entity 1: own vars + own state *)
     q2 := RS(q2, s2, r2);   (* entity 2: same code, other vars *)

   Key rules under current VeriSTC/VM semantics:
   1. FUNCTION bodies must be a single expression; the compiler
      inlines them at each call site (inline.v). Multi-statement
      bodies must be expanded by the upstream preprocessor.
   2. State variables (q1, q2) MUST be VAR_GLOBAL: the VM
      re-initializes PROGRAM frame locals to 0 every scan cycle,
      so locals cannot carry state across cycles. Globals live in
      the persistent MEM section.
   3. VAR_GLOBAL blocks must appear before the POU list.
   4. Multiple outputs: one return value per call. A second
      output is either derived at the call site (Q1 := NOT q) or
      provided by a sibling function sharing the same inputs.
   ================================================================ *)

VAR_GLOBAL
  q1 : BOOL;   (* RS entity 1 state/output *)
  q2 : BOOL;   (* RS entity 2 state/output *)
END_VAR

(* RS bistable: Q := S OR (Q_old AND NOT R); R has priority *)
FUNCTION RS : BOOL
VAR_INPUT
  Q_old : BOOL;
  S : BOOL;
  R : BOOL;
END_VAR
  RS := S OR (Q_old AND NOT R);
END_FUNCTION

PROGRAM MAIN
VAR
  s1 : BOOL;
  r1 : BOOL;
  s2 : BOOL;
  r2 : BOOL;
  tick : DINT;
END_VAR
  tick := CycleCounter();

  (* stimuli: entity 1 set@2 reset@6, entity 2 set@4 reset@8 *)
  s1 := tick = 2;
  r1 := tick = 6;
  s2 := tick = 4;
  r2 := tick = 8;

  (* multi-entity calls: original vars + previous state in,
     new state out via the single return value *)
  q1 := RS(q1, s1, r1);
  q2 := RS(q2, s2, r2);

  PRINT('tick', tick, q1, q2);
END_PROGRAM

(* ---- rs_multi_entity_fb.expanded.st ---- *)
(* ================================================================
   GENERATED by tools/stpreproc.py -- DO NOT EDIT BY HAND
   source: rs_multi_entity_fb.st
   template: rs_v1.tpl.st lib=demo version=1.2 sha256=39688997751b6fe4
   协议: PRE-1/2/5/7, T-1..T-4（实现一份: 共享函数实体）
   ================================================================ *)

VAR_GLOBAL
  fby1 : DINT;
END_VAR

FUNCTION FBY_RESET : DINT
VAR_INPUT
  fby   : DINT;
  reset : DINT;
END_VAR
  fby := reset;
  FBY_RESET := reset;
END_FUNCTION
(* @tpl RESET_END *)

(* @tpl FUNCTION *)
FUNCTION FBY : DINT
VAR_INPUT
  pre : DINT;
  q   : DINT;
END_VAR
  FBY := pre;
  pre := q;
END_FUNCTION

(* 实例声明：每个实体 = 同一模板的一份上下文 *)

PROGRAM MAIN
VAR
  tick  : DINT;
END_VAR
  tick := CycleCounter();
  IF tick = 1 THEN
    (* 初始化：调用共享函数实体，传入实例上下文 *)
    FBY_RESET(fby1, 0);
  END_IF;

  FBY(fby1, tick);

  (* 输出消费：读实例上下文全局（本 demo 只消费状态 Q） *)
  PRINT('tick=', tick, 'fby1=', fby1, '\n');
END_PROGRAM

(* ---- rs_multi_entity_fb.st ---- *)
(* ================================================================
   rs_multi_entity_fb.st  --  授权源文件（FB 形式多实体 RS）

   实现只在模板一份：lib-templates/rs_v1.tpl.st
   MAIN 只调用、不重新实现。编译器实际接收的是预处理展开产物：
     python3 tools/stpreproc.py \
       tests/st-examples/rs_multi_entity_fb.st \
       -o tests/st-examples/rs_multi_entity_fb.expanded.st
   （展开产物含生成头，标注模板版本与 sha256，见 PRE-5）

   与 FUNCTION 版 (rs_multi_entity.st) 的分工差异：
     FUNCTION 版: 状态由调用方搬进搬出   q1 := RS(q1, s1, r1);
     FB 版:      状态封装在实例上下文，MAIN 只见调用   rs1(S := ..., R := ...);
   ================================================================ *)

(* @use lib-templates/rs_v1.tpl.st *)

(* 实例声明：每个实体 = 同一模板的一份上下文 *)
(* @fb rs1 : RS_V1 *)
(* @fb rs2 : RS_V1 *)

PROGRAM MAIN
VAR
  tick  : DINT;
END_VAR
  tick := CycleCounter();

  (* 多实体调用：同一份模板实现，各绑各的输入 *)
  rs1(S := tick = 2, R := tick = 6);
  rs2(S := tick = 4, R := tick = 8);

  (* 输出消费：读实例上下文全局（本 demo 只消费状态 Q） *)
  PRINT('tick', tick, rs1.Q, rs2.Q);
END_PROGRAM
